		ELSE
				IF (_eDirection=E_Direction.DIRECTION_POSITIVE)THEN
					_fDistance:=_fPos-stAxis.stNcTOPLC.fActPos;
				ELSE
					_fDistance:=stAxis.stNcTOPLC.fActPos-_fPos;
				END_IF
		END_IF
		(*IF (_eDirection=E_Direction.DIRECTION_POSITIVE)THEN
			_fDistance:=_fPos-stAxis.stNcTOPLC.fActPos;
		ELSE
			_fDistance:=stAxis.stNcTOPLC.fActPos-_fPos;
		END_IF*)
		_nPathSegment:=1;
		_fAcc:=stAxis.stPLCTONC.stEndPosition.fAccleration;
	    _fDec:=stAxis.stPLCTONC.stEndPosition.fDeceleration;
ELSE
		_nPathSegment:=2;
		_fVeloStart:=stAxis.stNcTOPLC.fActVelo;
	    _fVeloEnd:=_fPreTaVel;
	    _fTargetVelo:=_fPreTaVel;
		_fDistance:=_fNewAccDis;
		_fAcc:=_fNewAcc;
	    _fDec:=_fNewAcc;
		_fPosIn:=_fDealt_S+_fPreDealt_S;       //11.29
	    _fVeloStart_2:=_fPreTaVel;
	    _fVeloEnd_2:=0.0;
	    _fTargetVelo_2:=_fPreTaVel;
		IF (stAxis.stPLCTONC.nRoadID_2<>0)AND (stAxis.stPLCTONC.nRoadID_1<>0)THEN   //判断指令
				IF (stAxis.stPLCTONC.stStartPosition.nRoadID<>stAxis.stPLCTONC.stEndPosition.nRoadID)THEN
				    IF(stAxis.stNcTOPLC.nCuRoadID=stAxis.stPLCTONC.nRoadID_2) THEN //第二路段
						IF (_eDirection=E_Direction.DIRECTION_POSITIVE)THEN
							 IF NOT stAxis.stPLCTONC.bRoadDirection  THEN   //正向 
								 _fDistance_2:=_fPos-stAxis.stPLCTONC.fRoad1_Length-stAxis.stNcTOPLC.fActPos-_fNewAccDis;
							 ELSE
								 _fDistance_2:=stAxis.stNcTOPLC.fActPos-(stAxis.stPLCTONC.fRoad2_Length-_fPos+stAxis.stPLCTONC.fRoad1_Length)-_fNewAccDis;
							 END_IF
						ELSE
							IF NOT stAxis.stPLCTONC.bRoadDirection  THEN   //正向 
								 _fDistance_2:=ABS(_fPos)-stAxis.stNcTOPLC.fActPos-_fNewAccDis;
							 ELSE
								 _fDistance_2:=stAxis.stNcTOPLC.fActPos-(stAxis.stPLCTONC.fRoad2_Length-ABS(_fPos))-_fNewAccDis;
							 END_IF
						END_IF
						stAxis.stPLCTONC.stStartPosition.nRoadID:=stAxis.stNcTOPLC.nCuRoadID;
					ELSE
						IF (_eDirection=E_Direction.DIRECTION_POSITIVE)THEN
							_fDistance_2:=_fPos-stAxis.stNcTOPLC.fActPos-_fNewAccDis;
						ELSE
							_fDistance_2:=stAxis.stNcTOPLC.fActPos-_fPos-_fNewAccDis;
						END_IF
					END_IF
				ELSE
					IF(stAxis.stNcTOPLC.nCuRoadID=stAxis.stPLCTONC.nRoadID_2) THEN //第二路段
						
						IF NOT stAxis.stPLCTONC.bRoadDirection  THEN   //正向 
							_fDistance_2:=_fPos-stAxis.stNcTOPLC.fActPos-_fNewAccDis;
						ELSE
							_fDistance_2:=stAxis.stNcTOPLC.fActPos-_fPos-_fNewAccDis;
						END_IF
						stAxis.stPLCTONC.stStartPosition.nRoadID:=stAxis.stNcTOPLC.nCuRoadID;
					ELSE
						IF (_eDirection=E_Direction.DIRECTION_POSITIVE)THEN
							_fDistance_2:=_fPos-stAxis.stNcTOPLC.fActPos-_fNewAccDis;
						ELSE
							_fDistance_2:=stAxis.stNcTOPLC.fActPos-_fPos-_fNewAccDis;
						END_IF
					END_IF
				END_IF
		ELSE
				IF (_eDirection=E_Direction.DIRECTION_POSITIVE)THEN
					_fDistance_2:=_fPos-stAxis.stNcTOPLC.fActPos-_fNewAccDis;
				ELSE
					_fDistance_2:=stAxis.stNcTOPLC.fActPos-_fPos-_fNewAccDis;
				END_IF
		END_IF
		(*IF (_eDirection=E_Direction.DIRECTION_POSITIVE)THEN
			_fDistance_2:=_fPos-stAxis.stNcTOPLC.fActPos-_fNewAccDis;
		ELSE
			_fDistance_2:=stAxis.stNcTOPLC.fActPos-_fPos-_fNewAccDis;
		END_IF*)
		_fAcc_2:=stAxis.stPLCTONC.stEndPosition.fAccleration;
	    _fDec_2:=stAxis.stPLCTONC.stEndPosition.fDeceleration;
		
END_IF
_bSynMode:=TRUE;
_bEnable:=TRUE;
stAxis.stAxisStatus.bSynDecActive:=TRUE;
IF GVL_MC.cDebug  THEN
	_sMessage:=FC_StrContact(stAxis,'next road dec2 gap control');
	 ADSLOGSTR(ADSLOG_MSGTYPE_HINT, _sMessage, '');
END_IF
END_ACTION

ACTION A_NextRoadGapControl:

//IF ((_fRealDis -_fGapSet)<=cDealtGap)AND(_pNextRoadPremover^.stAxisStatus.stPathRef.fTargetVelocity <stAxis.stAxisStatus.stPathRef.fTargetVelocity) THEN    //10.18 
(*IF ((_fRealDis -_fGapSet)<=_fSetDealtGap)AND(_pNextRoadPremover^.stAxisStatus.stPathRef.fTargetVelocity <stAxis.stAxisStatus.stPathRef.fTargetVelocity) THEN    //10.18
	
		_fPos:=stAxis.stPLCTONC.stEndPosition.fPosition;
		_fTargetVelo:=_pNextRoadPremover^.stAxisStatus.stPathRef.fTargetVelocity;
		_fVeloStart:=stAxis.stNcTOPLC.fActVelo;
		_fVeloEnd:=0;
		_fAcc:=stAxis.stPLCTONC.stEndPosition.fAccleration;
		_fDec:=stAxis.stPLCTONC.stEndPosition.fDeceleration;
		IF (_eDirection=E_Direction.DIRECTION_POSITIVE)THEN
		     _fDistance:=_fPos-stAxis.stNcTOPLC.fActPos;
	    ELSE
			 _fDistance:=stAxis.stNcTOPLC.fActPos-_fPos;
	    END_IF
		_bEnable:=TRUE;
		_nPathSegment:=1;
		stAxis.stAxisStatus.bSynDecActive:=TRUE;
		IF GVL_MC.cDebug  THEN
		     _sMessage:=FC_StrContact(stAxis,'nextroad gap control');
	         ADSLOGSTR(ADSLOG_MSGTYPE_HINT, _sMessage, '');
        END_IF
		RETURN;
END_IF *)

IF _fRealDis <=0 THEN   //05.19
	RETURN;
END_IF

IF (_pNextRoadPremover^.stAxisStatus.nNcCycleCounter<>0)THEN 
	 A_NextRoadCatchUp();
   // IF ((_fRealDis -_fGapSet)<=cDealtGap) THEN    //10.18 
	IF ((_fRealDis -_fGapSet)<=_fSetDealtGap) THEN    //10.18 	
			IF _fbDecNextPathTrig.Q THEN 
					   IF (stAxis.stPLCTONC.nRoadID_2<>0)AND (stAxis.stPLCTONC.nRoadID_1<>0)AND(stAxis.stNcTOPLC.nCuRoadID=stAxis.stPLCTONC.nRoadID_2)THEN
						   IF (stAxis.stPLCTONC.stStartPosition.nRoadID<>stAxis.stPLCTONC.stEndPosition.nRoadID)THEN
								IF (_eDirection=E_Direction.DIRECTION_POSITIVE)THEN
									IF NOT stAxis.stPLCTONC.bRoadDirection  THEN
										 _fPos:=stAxis.stPLCTONC.stEndPosition.fPosition-stAxis.stPLCTONC.fRoad1_Length;
									ELSE
										_fPos:=stAxis.stPLCTONC.fRoad2_Length-(stAxis.stPLCTONC.stEndPosition.fPosition-stAxis.stPLCTONC.fRoad1_Length);
									END_IF
									_fDistance:=ABS(stAxis.stNcTOPLC.fActPos-_fPos);
								ELSE
									IF NOT stAxis.stPLCTONC.bRoadDirection  THEN
										 _fPos:=ABS(stAxis.stPLCTONC.stEndPosition.fPosition);
									ELSE
										_fPos:=stAxis.stPLCTONC.fRoad2_Length-ABS(stAxis.stPLCTONC.stEndPosition.fPosition);
									END_IF
									_fDistance:=ABS(stAxis.stNcTOPLC.fActPos-_fPos);
								END_IF
						   ELSE
								_fPos:=stAxis.stPLCTONC.stEndPosition.fPosition;
								_fDistance:=ABS(stAxis.stNcTOPLC.fActPos-_fPos);
						   END_IF
					   ELSE
						   _fPos:=stAxis.stPLCTONC.stEndPosition.fPosition;
						   IF (_eDirection=E_Direction.DIRECTION_POSITIVE)THEN
							  _fDistance:=_fPos-stAxis.stNcTOPLC.fActPos;
						   ELSE
							  _fDistance:=stAxis.stNcTOPLC.fActPos-_fPos;
						   END_IF
					   END_IF
					   //_fPos:=stAxis.stPLCTONC.stEndPosition.fPosition;
					   IF _pNextRoadPremover^.stPLCTONC.bCmdDceUpdate THEN
							_fTargetVelo:=_pNextRoadPremover^.stPLCTONC.fTargetVelocity;
					   ELSE
						   _fTargetVelo:=_pNextRoadPremover^.stAxisStatus.stPathRef.fTargetVelocity;
					   END_IF
					   //_fTargetVelo:=_pNextRoadPremover^.stAxisStatus.stPathRef.fTargetVelocity;
					   _fVeloStart:=stAxis.stNcTOPLC.fActVelo;
					   _fVeloEnd:=0;
					   _fAcc:=stAxis.stPLCTONC.stEndPosition.fAccleration;
					   _fDec:=stAxis.stPLCTONC.stEndPosition.fDeceleration;
					   
					   _bEnable:=TRUE;
					   _nPathSegment:=1;
					   stAxis.stAxisStatus.bSynDecActive:=TRUE;
					   IF GVL_MC.cDebug  THEN
						_sMessage:=FC_StrContact(stAxis,'Nextroad SynDecActive path');
						 ADSLOGSTR(ADSLOG_MSGTYPE_HINT, _sMessage, '');
					   END_IF
			END_IF
	END_IF

END_IF
END_ACTION

ACTION A_NodeConfig:
IF stAxis.stNcTOPLC.nCuRoadID=0 THEN 
	RETURN;
END_IF 

_nMoverCounter:=GVL_MC.aRoadRef[stAxis.stNcTOPLC.nCuRoadID].nMoverCounter;
IF _nMoverCounter<>_nLastMoverCounter AND _nMoverCounter<>0  THEN 
	
    FOR _nNodeIndex:=1 TO GVL_MC.MAX_MOVER  DO
	    IF (GVL_MC.aRoadRef[stAxis.stNcTOPLC.nCuRoadID].aNode[_nNodeIndex].nAxisId=stAxis.stNcTOPLC.nAxisId)THEN
			stAxis.stAxisStatus.pPremover:=GVL_MC.aRoadRef[stAxis.stNcTOPLC.nCuRoadID].aNode[_nNodeIndex].pPremover;
	        stAxis.stAxisStatus.pAftermover:=GVL_MC.aRoadRef[stAxis.stNcTOPLC.nCuRoadID].aNode[_nNodeIndex].pAftermover;
			EXIT;
		END_IF
   END_FOR
   _nLastMoverCounter:=GVL_MC.aRoadRef[stAxis.stNcTOPLC.nCuRoadID].nMoverCounter;   //05.08 修改前置后置更新条件
END_IF
END_ACTION

ACTION A_NodeUpdate:
// road node 更新
// 动子出现在某road上增加 01.09
_fbTrigRoadUpdate(CLK:=stAxis.stCodToNCParam.bArrayReseved1 , Q=> );
//IF stAxis.stNcTOPLC.nCuRoadID=0 AND stAxis.stCodToNCParam.bArrayReseved1  AND stAxis.stCodToNCParam.nRoadID<>0 THEN
IF _fbTrigRoadUpdate.Q  AND stAxis.stCodToNCParam.nRoadID<>0 AND NOT _bInsertOk THEN
	stAxis.stNcTOPLC.nCuRoadID:=stAxis.stCodToNCParam.nRoadID;
	_bInsertOk :=_fbAxisGroupList.M_InsertNode(aRoadRef:=GVL_MC.aRoadRef , nSysType:=stAxis.stAxisParam.stRoadParam.nSysType , nRoadId:=stAxis.stCodToNCParam.nRoadID , pAixs:=ADR(stAxis) );
    (*IF GVL_MC.cDebug  THEN
	    _sMessage2:=FC_StrContactEx(stAxis,'insertAxis');
	     ADSLOGSTR(ADSLOG_MSGTYPE_HINT, _sMessage2, '');
    END_IF*)
	_sMessage3:='';
	_sMessage3:=CONCAT(DWORD_TO_STRING(stAxis.stNcTOPLC.nAxisId),',insertAxis');
	IF stAxis.stNcTOPLC.nCuRoadID>0 AND stAxis.stNcTOPLC.nCuRoadID<=GVL_MC.cRoadNum AND GVL_MC.cDebug THEN
		IF GVL_MC.aRoadRef[stAxis.stNcTOPLC.nCuRoadID].nMoverCounter>0  THEN
			FOR _nPreIndex:=1 TO GVL_MC.aRoadRef[stAxis.stNcTOPLC.nCuRoadID].nMoverCounter   DO
				_sMessage3:=CONCAT(_sMessage3,DWORD_TO_STRING(GVL_MC.aRoadRef[stAxis.stNcTOPLC.nCuRoadID].aNode[_nPreIndex].nAxisId));
				_sMessage3:=CONCAT(_sMessage3,',');
			END_FOR
			ADSLOGSTR(ADSLOG_MSGTYPE_HINT, _sMessage3, '');
		END_IF
	END_IF
END_IF
IF NOT stAxis.stCodToNCParam.bArrayReseved1 THEN
	_bInsertOk:=FALSE;
END_IF
// 07.04
IF stAxis.stNcTOPLC.nCuRoadID=0 THEN 
	RETURN;
END_IF 

_fbTrigRoadDeleUpdate(CLK:=stAxis.stCodToNCParam.bArrayReseved2 , Q=> );   //01.29
IF _fbTrigRoadDeleUpdate.Q THEN
	_bDeleteNodeOk:=_fbAxisGroupList.M_DeleteNode(aRoadRef:=GVL_MC.aRoadRef , nSysType:=stAxis.stAxisParam.stRoadParam.nSysType , nRoadId:=stAxis.stNcTOPLC.nCuRoadID , pAixs:=ADR(stAxis));
	(*IF GVL_MC.cDebug  THEN
	    _sMessage2:=FC_StrContactEx(stAxis,'deleteAxis');
	     ADSLOGSTR(ADSLOG_MSGTYPE_HINT, _sMessage2, '');
    END_IF*)
	_sMessage3:='';
	_sMessage3:=CONCAT(DWORD_TO_STRING(stAxis.stNcTOPLC.nAxisId),',deleteAxis');
    IF stAxis.stNcTOPLC.nCuRoadID>0 AND stAxis.stNcTOPLC.nCuRoadID<=GVL_MC.cRoadNum AND GVL_MC.cDebug THEN
	    IF GVL_MC.aRoadRef[stAxis.stNcTOPLC.nCuRoadID].nMoverCounter>0 THEN
			FOR _nPreIndex:=1 TO GVL_MC.aRoadRef[stAxis.stNcTOPLC.nCuRoadID].nMoverCounter   DO
				_sMessage3:=CONCAT(_sMessage3,DWORD_TO_STRING(GVL_MC.aRoadRef[stAxis.stNcTOPLC.nCuRoadID].aNode[_nPreIndex].nAxisId));
				_sMessage3:=CONCAT(_sMessage3,',');
			END_FOR
			ADSLOGSTR(ADSLOG_MSGTYPE_HINT, _sMessage3, '');
		END_IF
	END_IF
END_IF

// 先增加后删除
(*IF stAxis.stNcTOPLC.nCuRoadID=0 THEN 
	RETURN;
END_IF *) //07.04
IF (_nLastRoadID<>stAxis.stNcTOPLC.nCuRoadID) AND (_nLastRoadID<>0)THEN
	
	_nLastMoverCounter:=GVL_MC.aRoadRef[stAxis.stNcTOPLC.nCuRoadID].nMoverCounter;  //********重新修改前置后质更新条件     05.08
	_bAddNodeOk :=_fbAxisGroupList.M_AddNode(aRoadRef:=GVL_MC.aRoadRef , nRoadId:=stAxis.stNcTOPLC.nCuRoadID , pAixs:=ADR(stAxis));
	//_bAddNodeOk :=_fbAxisGroupList.M_InsertNode(aRoadRef:=GVL_MC.aRoadRef , nSysType:=stAxis.stAxisParam.stRoadParam.nSysType , nRoadId:=stAxis.stNcTOPLC.nCuRoadID , pAixs:=ADR(stAxis) );
    _bDeleteNodeOk:=_fbAxisGroupList.M_DeleteNode(aRoadRef:=GVL_MC.aRoadRef , nSysType:=stAxis.stAxisParam.stRoadParam.nSysType , nRoadId:=_nLastRoadID , pAixs:=ADR(stAxis));
	(*IF GVL_MC.cDebug  THEN
	    //_sMessage2:=FC_StrContactEx(stAxis,'roadchange');
	    // ADSLOGSTR(ADSLOG_MSGTYPE_HINT, _sMessage2, '');
		  _sMessage3:=CONCAT(DWORD_TO_STRING(stAxis.stNcTOPLC.nAxisId),',roadchange');
		  _sMessage3:=CONCAT(_sMessage3,',');
		  _sMessage3:=CONCAT(_sMessage3,LREAL_TO_STRING(stAxis.stNcTOPLC.fActPos));
		  _sMessage3:=CONCAT(_sMessage3,',');
		  _sMessage3:=CONCAT(_sMessage3,DWORD_TO_STRING(GVL_MC.aRoadRef[stAxis.stNcTOPLC.nCuRoadID].aNode[GVL_MC.aRoadRef[stAxis.stNcTOPLC.nCuRoadID].nMoverCounter].pMover^.stNcTOPLC.nAxisId));
          _sMessage3:=CONCAT(_sMessage3,',');	 
		  _sMessage3:=CONCAT(_sMessage3,LREAL_TO_STRING(GVL_MC.aRoadRef[stAxis.stNcTOPLC.nCuRoadID].aNode[GVL_MC.aRoadRef[stAxis.stNcTOPLC.nCuRoadID].nMoverCounter].pMover^.stNcTOPLC.fActPos));
   	      _sMessage3:=CONCAT(_sMessage3,',');
		  _sMessage3:=CONCAT(_sMessage3,UINT_TO_STRING(GVL_MC.aRoadRef[stAxis.stNcTOPLC.nCuRoadID].nMoverCounter));
		  ADSLOGSTR(ADSLOG_MSGTYPE_HINT, _sMessage3, '');
    END_IF*)
	_sMessage3:='';
	_sMessage3:=CONCAT(DWORD_TO_STRING(stAxis.stNcTOPLC.nAxisId),',roadchange');
	IF stAxis.stNcTOPLC.nCuRoadID>0 AND stAxis.stNcTOPLC.nCuRoadID<=GVL_MC.cRoadNum AND GVL_MC.cDebug THEN
		IF GVL_MC.aRoadRef[stAxis.stNcTOPLC.nCuRoadID].nMoverCounter>0  THEN
			FOR _nPreIndex:=1 TO GVL_MC.aRoadRef[stAxis.stNcTOPLC.nCuRoadID].nMoverCounter   DO
				
				_sMessage3:=CONCAT(_sMessage3,DWORD_TO_STRING(GVL_MC.aRoadRef[stAxis.stNcTOPLC.nCuRoadID].aNode[_nPreIndex].nAxisId));
				_sMessage3:=CONCAT(_sMessage3,',');
			END_FOR
			ADSLOGSTR(ADSLOG_MSGTYPE_HINT, _sMessage3, '');
		END_IF
	END_IF
END_IF



_nLastRoadID:=stAxis.stNcTOPLC.nCuRoadID;

_bAddNodeOk:=FALSE;
_bDeleteNodeOk:=FALSE;
END_ACTION

ACTION A_Planning:
IF (stAxis.stPLCTONC.ePlanningMode=E_PlanningMode.PLANNINGMODE_TSHAPED)THEN 
   A_TShaped();
ELSIF (stAxis.stPLCTONC.ePlanningMode=E_PlanningMode.PLANNINGMODE_SSHAPED)THEN 
   A_SShapedPlanning();
ELSIF (stAxis.stPLCTONC.ePlanningMode=E_PlanningMode.PLANNINGMODE_LINEAR)THEN 
  A_LinearPlanning();

ELSIF (stAxis.stPLCTONC.ePlanningMode=E_PlanningMode.PLANNINGMODE_FOLLOWMASTER)THEN 
  A_FollowMasterPlanning();
  
ELSIF (stAxis.stPLCTONC.ePlanningMode=E_PlanningMode.PLANNINGMODE_PLOYNOM3)THEN 
	A_Ploynom3Planning();
ELSIF (stAxis.stPLCTONC.ePlanningMode=E_PlanningMode.PLANNINGMODE_FOLLOW)THEN 
	A_FollowPlanning();	
ELSE 
   A_TShaped();

END_IF
END_ACTION

ACTION A_Ploynom3Planning:
//_fbAxis.strStartPoint.fPosition:=stAxis.stNcTOPLC.fActPos;
//_fbAxis.strEndPoint.fPosition:=stAxis.stPLCTONC.stEndPosition.fPosition;
_fbAxis.strStartPoint.fPosition:=0;
_fbAxis.strEndPoint.fPosition:=ABS(stAxis.stPLCTONC.stEndPosition.fPosition-stAxis.stNcTOPLC.fActPos)/ABS(stAxis.stPLCTONC.stMasterParam.fEndPos-stAxis.stPLCTONC.stMasterParam.fStartPos);

IF (stAxis.stAxisStatus.pMaster^.stNcTOPLC.fActVelo<>0)  THEN 
    _fbAxis.strStartPoint.fVelocity :=stAxis.stNcTOPLC.fActVelo/stAxis.stAxisStatus.pMaster^.stNcTOPLC.fActVelo;
ELSE
	_fbAxis.strStartPoint.fVelocity :=0;
END_IF

//_fbAxis.strEndPoint.fVelocity:=stAxis.stAxisStatus.stPathRef.fVeloRatio;
_fbAxis.strEndPoint.fVelocity:=stAxis.stPLCTONC.fGearRatio;
_stPolynom5Factor:=_fbAxis.M_Ploynom3(fTheat_Start:=0 ,
               fTheat_End:=1  );
			   

_bCalculateDone:=TRUE;
END_ACTION

ACTION A_Ploynom3Position:
_nSysType:=stAxis.stPLCTONC.nSysType;
stAxis.stNcTOPLC.nAxisState:=6;
stAxis.stAxisStatus.nNcCycleCounter:=stAxis.stAxisStatus.nNcCycleCounter+1;
_fMasterStartPos:=stAxis.stPLCTONC.stMasterParam.fStartPos;
_fMasterEndPos:=stAxis.stPLCTONC.stMasterParam.fEndPos;

_fSlaveStartPos:=stAxis.stPLCTONC.stStartPosition.fPosition;
// 自变量区间归一化

_fDealt_X:=ABS(_fMasterEndPos-_fMasterStartPos);
IF (_fDealt_X<=0)THEN 
	RETURN;
END_IF
_fPos_X:=ABS(stAxis.stAxisStatus.pMaster^.stNcTOPLC.fActPos-_fMasterStartPos)/_fDealt_X;

IF (_fPos_X<=1)THEN

	// 归一化从轴位置、速度、加速度和加加速计算
	_stAxis_Point.fPosition:=_stPolynom5Factor.fA0+ _stPolynom5Factor.fA1*_fPos_X+ _stPolynom5Factor.fA2*_fPos_X*_fPos_X
						   +_stPolynom5Factor.fA3*_fPos_X*_fPos_X*_fPos_X; 
						   
	_stAxis_Point.fVelocity:=_stPolynom5Factor.fA1+ 2*_stPolynom5Factor.fA2*_fPos_X+3*_stPolynom5Factor.fA3*_fPos_X*_fPos_X;
	
	_stAxis_Point.fAccleration:=2*_stPolynom5Factor.fA2+6*_stPolynom5Factor.fA3*_fPos_X;
	_stAxis_Point.fbJerk:=6*_stPolynom5Factor.fA3;
	
	IF stAxis.stAxisStatus.bPositiveDirection THEN
		stAxis.stNcTOPLC.fActPos:=_fDealt_X*_stAxis_Point.fPosition+_fSlaveStartPos;    
	ELSE
		stAxis.stNcTOPLC.fActPos:=_fSlaveStartPos-_fDealt_X*_stAxis_Point.fPosition;    
	END_IF                  
	stAxis.stNcTOPLC.fSetVelo:=_stAxis_Point.fVelocity*ABS(stAxis.stAxisStatus.pMaster^.stNcTOPLC.fActVelo);
	stAxis.stNcTOPLC.fSetAcc:=_stAxis_Point.fAccleration*ABS(stAxis.stAxisStatus.pMaster^.stNcTOPLC.fActVelo*stAxis.stAxisStatus.pMaster^.stNcTOPLC.fActVelo)/_fDealt_X;
	stAxis.stNcTOPLC.fSetJerk:=_stAxis_Point.fbJerk*ABS(stAxis.stAxisStatus.pMaster^.stNcTOPLC.fActVelo*stAxis.stAxisStatus.pMaster^.stNcTOPLC.fActVelo*stAxis.stAxisStatus.pMaster^.stNcTOPLC.fActVelo)/(_fDealt_X*_fDealt_X);
							  
	stAxis.stNcTOPLC.fActVelo:=stAxis.stNcTOPLC.fSetVelo;
	_stAxis_Point.fPosition:=stAxis.stNcTOPLC.fActPos;
ELSE
	stAxis.stNcTOPLC.fSetVelo:=LTRUNC(stAxis.stAxisStatus.pMaster^.stNcTOPLC.fActVelo*stAxis.stPLCTONC.fGearRatio);
    stAxis.stNcTOPLC.fActVelo:=LTRUNC(stAxis.stAxisStatus.pMaster^.stNcTOPLC.fActVelo*stAxis.stPLCTONC.fGearRatio);
    IF stAxis.stAxisStatus.bPositiveDirection THEN
         _stAxis_Point.fPosition:=stAxis.stAxisStatus.pMaster^.stNcTOPLC.fDealtPos*stAxis.stPLCTONC.fGearRatio +_stAxis_Point.fPosition;

    ELSE
        _stAxis_Point.fPosition:=-stAxis.stAxisStatus.pMaster^.stNcTOPLC.fDealtPos*stAxis.stPLCTONC.fGearRatio +_stAxis_Point.fPosition;
    END_IF
	stAxis.stNcTOPLC.fDealtPos:=ABS(LTRUNC(_stAxis_Point.fPosition)-stAxis.stNcTOPLC.fActPos);    //01.13
	stAxis.stNcTOPLC.fActPos:=LTRUNC(_stAxis_Point.fPosition);
END_IF
END_ACTION

ACTION A_Ploynom5Position:
_bEndOfProfile:=FALSE;
_nSysType:=stAxis.stPLCTONC.nSysType;
stAxis.stNcTOPLC.nAxisState:=6;
stAxis.stAxisStatus.nNcCycleCounter:=stAxis.stAxisStatus.nNcCycleCounter+1;

//数据装载
IF stAxis.stPLCTONC.stCamParam.bCamLoad THEN 
   _stCamParam:=stAxis.stPLCTONC.stCamParam;
   stAxis.stPLCTONC.stCamParam.bCamLoad:=FALSE;
END_IF 

//buffer 更新
 _fbCamBufUpdateTrig(CLK:= (INT_TO_UINT(_nIndex)=(cPointBuffer-1)OR (NOT _bFisrtUpdate)), Q=> );

IF(_stCamParam.nElements> cPointBuffer) THEN
   IF _fbCamBufUpdateTrig.Q   THEN
      _aCamBuffer:=_stCamParam.aCamBuffer;
	  _nIndex:=0;
	  _nCamBufferNum:=_nCamBufferNum+1;
   END_IF 
ELSE
	_aCamBuffer:=_stCamParam.aCamBuffer;
	_nCamBufferNum:=1;
END_IF

// 点更新及曲线系数计算
_fbCamPointUpdateTrig(CLK:=(_nIndex<>_nLastIndex)OR (NOT _bFisrtUpdate)   , Q=> );
IF _fbCamPointUpdateTrig.Q THEN
     IF (_stCamParam.nPointType=1) THEN  //xyva
         _fMasterStartPos:=_aCamBuffer[_nIndex].fDx;
	     _fMasterEndPos:=_aCamBuffer[_nIndex+1].fDx;
	     _fDealt_X:=ABS(_fMasterEndPos-_fMasterStartPos);
		 IF (_fDealt_X=0)THEN 
			 RETURN;
		 END_IF
		_fSlaveStartPos :=_aCamBuffer[_nIndex].fDy;
		_fbAxis.strStartPoint.fPosition:=0;
		_fbAxis.strEndPoint.fPosition:=ABS((_aCamBuffer[_nIndex+1].fDy-_fSlaveStartPos))/_fDealt_X;
		_fbAxis.strStartPoint.fVelocity :=_aCamBuffer[_nIndex].fDv;
		_fbAxis.strEndPoint.fVelocity:=_aCamBuffer[_nIndex+1].fDv;
		_fbAxis.strStartPoint.fAccleration :=_aCamBuffer[_nIndex].fDa*_fDealt_X;
		_fbAxis.strEndPoint.fAccleration:=_aCamBuffer[_nIndex+1].fDa*_fDealt_X;
		_fbAxis.strStartPoint.fbJerk :=_aCamBuffer[_nIndex].fDa*_fDealt_X*_fDealt_X;
		_fbAxis.strEndPoint.fbJerk:=_aCamBuffer[_nIndex+1].fDa*_fDealt_X*_fDealt_X;
	 ELSIF (_stCamParam.nPointType=2) THEN   //xy
		 _fMasterStartPos:=_aCamBuffer[_nIndex].fDx;
	     _fMasterEndPos:=_aCamBuffer[_nIndex+1].fDx;
	     _fDealt_X:=ABS(_fMasterEndPos-_fMasterStartPos);
		 _fSlaveStartPos :=_aCamBuffer[_nIndex].fDy;
		 _fbAxis.strStartPoint.fPosition:=0;
		 IF (_fDealt_X=0)THEN 
			 RETURN;
		 END_IF
		 _fbAxis.strEndPoint.fPosition:=ABS(_aCamBuffer[_nIndex+1].fDy-_fSlaveStartPos)/_fDealt_X;
		 IF (_nIndex=0)AND (_nCamBufferNum=1)THEN
		    _fbAxis.strStartPoint.fVelocity :=0;
			_fbAxis.strStartPoint.fAccleration :=0;
		 ELSE
			 _fbAxis.strStartPoint.fVelocity :=1;
			 _fbAxis.strStartPoint.fAccleration :=0;
		 END_IF

		 _fbAxis.strEndPoint.fVelocity:=1;
		 IF _stCamParam.bPeriodic AND (stAxis.stNcTOPLC.nCuSegIndex =(_stCamParam.nElements-1)) THEN
			 _fbAxis.strEndPoint.fVelocity:=0;
		 END_IF
		 _fbAxis.strStartPoint.fAccleration :=0;
		 _fbAxis.strEndPoint.fAccleration:=0;
		 _fbAxis.strStartPoint.fbJerk :=0;
		 _fbAxis.strEndPoint.fbJerk:=0;
		
     ELSE
		 RETURN;
		 
	 END_IF
	_stPolynom5Factor:=_fbAxis.M_Ploynom5(fTheat_Start:=0 ,fTheat_End:=1);
	_bFisrtUpdate:=TRUE;
END_IF 
_nLastIndex :=_nIndex;
IF (_fDealt_X=0)THEN 
	RETURN;
END_IF
// 位置计算

// 自变量区间归一化
//_fDealt_X:=_fMasterEndPos-_fMasterStartPos;
IF stAxis.stAxisStatus.bPositiveDirection  THEN
    _fPos_X:=(stAxis.stAxisStatus.pMaster^.stNcTOPLC.fActPos-_fMasterStartPos)/ABS(_fDealt_X);
ELSE
	_fPos_X:=(_fMasterStartPos-stAxis.stAxisStatus.pMaster^.stNcTOPLC.fActPos)/ABS(_fDealt_X);
END_IF

IF (_fPos_X<0)THEN 
	RETURN;
END_IF

_stAxis_Point.fPosition:=_stPolynom5Factor.fA0+ _stPolynom5Factor.fA1*_fPos_X+ _stPolynom5Factor.fA2*_fPos_X*_fPos_X
                        +_stPolynom5Factor.fA3*_fPos_X*_fPos_X*_fPos_X+_stPolynom5Factor.fA4*_fPos_X*_fPos_X*_fPos_X*_fPos_X
						+_stPolynom5Factor.fA5*_fPos_X*_fPos_X*_fPos_X*_fPos_X*_fPos_X;
                          
						
_stAxis_Point.fVelocity:=_stPolynom5Factor.fA1+ 2*_stPolynom5Factor.fA2*_fPos_X+3*_stPolynom5Factor.fA3*_fPos_X*_fPos_X
                          +4*_stPolynom5Factor.fA4*_fPos_X*_fPos_X*_fPos_X+5*_stPolynom5Factor.fA5*_fPos_X*_fPos_X*_fPos_X*_fPos_X;
                          
_stAxis_Point.fAccleration:= 2*_stPolynom5Factor.fA2+6*_stPolynom5Factor.fA3*_fPos_X+12*_stPolynom5Factor.fA4*_fPos_X*_fPos_X+20*_stPolynom5Factor.fA5*_fPos_X*_fPos_X*_fPos_X;
_stAxis_Point.fbJerk:=6*_stPolynom5Factor.fA3+24*_stPolynom5Factor.fA4*_fPos_X+60*_stPolynom5Factor.fA5*_fPos_X*_fPos_X;

IF stAxis.stAxisStatus.bPositiveDirection THEN 
	//stAxis.stNcTOPLC.fSetPos:=_stAxis_Point.fPosition*_fDealt_X+_fSlaveStartPos;
	stAxis.stNcTOPLC.fActPos:=_stAxis_Point.fPosition*_fDealt_X+_fSlaveStartPos;
	stAxis.stNcTOPLC.fSetVelo:=_stAxis_Point.fVelocity*ABS(stAxis.stAxisStatus.pMaster^.stNcTOPLC.fActVelo);
	stAxis.stNcTOPLC.fSetAcc:=_stAxis_Point.fAccleration*ABS(stAxis.stAxisStatus.pMaster^.stNcTOPLC.fActVelo*stAxis.stAxisStatus.pMaster^.stNcTOPLC.fActVelo)/_fDealt_X;
	stAxis.stNcTOPLC.fSetJerk:=_stAxis_Point.fbJerk*ABS(stAxis.stAxisStatus.pMaster^.stNcTOPLC.fActVelo*stAxis.stAxisStatus.pMaster^.stNcTOPLC.fActVelo*stAxis.stAxisStatus.pMaster^.stNcTOPLC.fActVelo)/(_fDealt_X*_fDealt_X);
	//stAxis.stNcTOPLC.fActPos:=stAxis.stNcTOPLC.fSetPos;
	stAxis.stNcTOPLC.fActVelo:=stAxis.stNcTOPLC.fSetVelo;
ELSE
	//stAxis.stNcTOPLC.fSetPos:=-_stAxis_Point.fPosition*_fDealt_X+_fSlaveStartPos;
	stAxis.stNcTOPLC.fActPos:=-_stAxis_Point.fPosition*_fDealt_X+_fSlaveStartPos;
	stAxis.stNcTOPLC.fSetVelo:=_stAxis_Point.fVelocity*ABS(stAxis.stAxisStatus.pMaster^.stNcTOPLC.fActVelo);
	stAxis.stNcTOPLC.fSetAcc:=_stAxis_Point.fAccleration*ABS(stAxis.stAxisStatus.pMaster^.stNcTOPLC.fActVelo*stAxis.stAxisStatus.pMaster^.stNcTOPLC.fActVelo)/_fDealt_X;
	stAxis.stNcTOPLC.fSetJerk:=_stAxis_Point.fbJerk*ABS(stAxis.stAxisStatus.pMaster^.stNcTOPLC.fActVelo*stAxis.stAxisStatus.pMaster^.stNcTOPLC.fActVelo*stAxis.stAxisStatus.pMaster^.stNcTOPLC.fActVelo)/(_fDealt_X*_fDealt_X);
	//stAxis.stNcTOPLC.fActPos:=stAxis.stNcTOPLC.fSetPos;
	stAxis.stNcTOPLC.fActVelo:=stAxis.stNcTOPLC.fSetVelo;
END_IF
(*IF (_nSysType=3)THEN   //环形
	IF stAxis.stAxisStatus.bPositiveDirection THEN
		stAxis.stNcTOPLC.nModuloSetTurns:=LREAL_TO_DINT(LTRUNC(stAxis.stNcTOPLC.fSetPos/stAxis.stNcTOPLC.fModuloFactor));
	ELSE
		IF stAxis.stNcTOPLC.fSetPos<(stAxis.stNcTOPLC.nModuloSetTurns*stAxis.stNcTOPLC.fModuloFactor)THEN 
				stAxis.stNcTOPLC.nModuloSetTurns:=stAxis.stNcTOPLC.nModuloSetTurns-1;
		END_IF
	END_IF
	stAxis.stNcTOPLC.fModuloSetPos:= MODABS(stAxis.stNcTOPLC.fSetPos,stAxis.stNcTOPLC.fModuloFactor);
ELSE
	stAxis.stNcTOPLC.fModuloSetPos:= ABS(stAxis.stNcTOPLC.fSetPos);
END_IF*)


stAxis.stNcTOPLC.nCuSegIndex:=INT_TO_UINT(_nIndex+1)+(_nCamBufferNum-1)*cPointBuffer;
// index更新
IF stAxis.stAxisStatus.bPositiveDirection THEN 
	IF (stAxis.stNcTOPLC.fActPos>=_aCamBuffer[_nIndex+1].fDy)THEN 
		_nIndex:=_nIndex+1;
		IF stAxis.stNcTOPLC.nCuSegIndex >(_stCamParam.nElements-1) THEN      //结束条件判断
			_bCalculateDone:=FALSE;
			_nIndex:=0;
			_nLastIndex :=0;
			 stAxis.stAxisStatus.stPathRef.bCalculateDone:=FALSE;
			 stAxis.stNcTOPLC.nAxisState:=2;
		 
			 stAxis.stNcTOPLC.fSetAcc:=0;
			 _bFisrtUpdate:=FALSE;
			 stAxis.stNcTOPLC.nCuSegIndex:=0;
			 _nCamBufferNum:=0;
			 _fDealt_X:=0;
			 _fbCamBufUpdateTrig(CLK:= FALSE, Q=> );
			 _fbCamPointUpdateTrig(CLK:=FALSE   , Q=> );
			 _bEndOfProfile:=TRUE;
		END_IF
	END_IF
ELSE
	IF (stAxis.stNcTOPLC.fActPos<=_aCamBuffer[_nIndex+1].fDy)THEN 
		_nIndex:=_nIndex+1;
		IF stAxis.stNcTOPLC.nCuSegIndex >(_stCamParam.nElements-1) THEN      //结束条件判断
			_bCalculateDone:=FALSE;
			_nIndex:=0;
			_nLastIndex :=0;
			 stAxis.stAxisStatus.stPathRef.bCalculateDone:=FALSE;
			 stAxis.stNcTOPLC.nAxisState:=2;
		 
			 stAxis.stNcTOPLC.fSetAcc:=0;
			 _bFisrtUpdate:=FALSE;
			 stAxis.stNcTOPLC.nCuSegIndex:=0;
			 _nCamBufferNum:=0;
			 _fDealt_X:=0;
			 _fbCamBufUpdateTrig(CLK:= FALSE, Q=> );
			 _fbCamPointUpdateTrig(CLK:=FALSE   , Q=> );
			 _bEndOfProfile:=TRUE;
		END_IF
	END_IF
END_IF
END_ACTION

ACTION A_PositionHandle:
//stAxis.stNcTOPLC.fActPos 输入
//stAxis.stNcTOPLC.fSetPos输出
IF (stAxis.stPLCTONC.eCommand=E_Command.COMMAND_ABSOLUTEFORK)OR (stAxis.stPLCTONC.eCommand=E_Command.COMMAND_CAMIN)OR 
	(stAxis.stPLCTONC.eCommand=E_Command.COMMAND_GEARINPOS)THEN
	stAxis.stNcTOPLC.fSetPos:=stAxis.stNcTOPLC.fActPos;
    
ELSE
	IF (stAxis.stAxisParam.stRoadParam.nSysType=1) OR (stAxis.stAxisParam.stRoadParam.nSysType=4) THEN 
		stAxis.stNcTOPLC.fSetPos:=stAxis.stNcTOPLC.fActPos;
	ELSE
		_fbFilterV2(nWindowSize:=nWindowSize , fData:=stAxis.stNcTOPLC.fActPos , fOutputData=>stAxis.stNcTOPLC.fSetPos );
	END_IF
END_IF

IF (stAxis.stPLCTONC.nSysType=3)THEN
	IF stAxis.stAxisStatus.bPositiveDirection THEN
		stAxis.stNcTOPLC.nModuloSetTurns:=LREAL_TO_DINT(LTRUNC(stAxis.stNcTOPLC.fActPos/stAxis.stNcTOPLC.fModuloFactor));
	ELSE
		IF stAxis.stNcTOPLC.fActPos<(stAxis.stNcTOPLC.nModuloSetTurns*stAxis.stNcTOPLC.fModuloFactor)THEN 
			 stAxis.stNcTOPLC.nModuloSetTurns:=stAxis.stNcTOPLC.nModuloSetTurns-1;
		END_IF
	END_IF
							
	stAxis.stNcTOPLC.fModuloSetPos:= MODABS(stAxis.stNcTOPLC.fSetPos,stAxis.stNcTOPLC.fModuloFactor);
ELSE
	stAxis.stNcTOPLC.fModuloSetPos:=ABS(stAxis.stNcTOPLC.fSetPos);
	// 04.30增加环形位置同步
	IF (stAxis.stAxisParam.stRoadParam.nSysType=3)THEN
		stAxis.stNcTOPLC.fModuloSetPos:= MODABS(stAxis.stNcTOPLC.fSetPos,stAxis.stNcTOPLC.fModuloFactor);
	END_IF
END_IF
END_ACTION

ACTION A_SShapedPlanning:
_stSShapedParam:=_fbAxis.M_SShaped(
					fStartPos:=_fStartPos , 
					fEndPos:=_fEndPos , 
					fStartVelo:=_fVeloStart , 
					fEndVelo:=_fVeloEnd , 
					fTargetVelo:=_fTargetVelo , 
					fTargetAcc:=_fAcc , 
					fTargetJerk:=_fJerk );
					
_stPathRef._nPathSegmentNum:=1;
_stPathRef.aExecutablePath[0].fTa:=_stSShapedParam.fTa;
_stPathRef.aExecutablePath[0].fTv:=_stSShapedParam.fTv;
_stPathRef.aExecutablePath[0].fTd:=_stSShapedParam.fTd;
_stPathRef.aExecutablePath[0].fTj1:=_stSShapedParam.fTj1;
_stPathRef.aExecutablePath[0].fTj2:=_stSShapedParam.fTj2;
_stPathRef.aExecutablePath[0].fTotalTime:=_stSShapedParam.fT;


_stPathRef.aExecutablePath[0].fStartVelo:=_fVeloStart;
_stPathRef.aExecutablePath[0].fExpVelo:=_stSShapedParam.fVlim;
_stPathRef.aExecutablePath[0].fEndVelo:=_fVeloEnd;
_stPathRef.aExecutablePath[0].fAccleration:=_stSShapedParam.fA_LimAcc ;
_stPathRef.aExecutablePath[0].fDeceleration:=_stSShapedParam.fA_LimDec;

_stPathRef.aExecutablePath[0].fJmax:=_stSShapedParam.fJmax ;
_stPathRef.aExecutablePath[0].fJmin:=_stSShapedParam.fJmin ;

_stPathRef.aExecutablePath[0].fStartPos:=_fStartPos;
_stPathRef.aExecutablePath[0].fEndPos:=_fEndPos;


_stPathRef.bCalculateDone:=TRUE;
stAxis.stAxisStatus.stPathRef:=_stPathRef;
_bCalculateDone:=TRUE;
_fTime:=0;
_nIndex:=0;
stAxis.stAxisStatus.nNcCycleCounter:=0;
END_ACTION

ACTION A_SShapedPosition:
stAxis.stNcTOPLC.nAxisState:=6;
_fTime:=_fTime+fCycleTime;
stAxis.stAxisStatus.nNcCycleCounter:=stAxis.stAxisStatus.nNcCycleCounter+1;


_stAxis_Point:=_fbAxis.M_SShapedPosition(fTime:=_fTime , stS_Parameter:=_stSShapedParam )	;					

//stAxis.stNcTOPLC.fSetPos:=_stAxis_Point.fPosition;
//stAxis.stNcTOPLC.fActPos:=stAxis.stNcTOPLC.fSetPos;
stAxis.stNcTOPLC.fActPos:=_stAxis_Point.fPosition;		
//stAxis.stNcTOPLC.fSetVelo:=_stAxis_Point.fVelocity;  //04.15注释
stAxis.stNcTOPLC.fActVelo:=_stAxis_Point.fVelocity;

IF (_eDirection=E_Direction.DIRECTION_POSITIVE)THEN    //04.15速度方向处理
	 stAxis.stNcTOPLC.fSetVelo:=stAxis.stNcTOPLC.fActVelo;
ELSE
     stAxis.stNcTOPLC.fSetVelo:=-stAxis.stNcTOPLC.fActVelo;
END_IF
	
stAxis.stNcTOPLC.fSetAcc:=_stAxis_Point.fAccleration;  //07.30
stAxis.stNcTOPLC.fSetJerk:=_stAxis_Point.fbJerk;

//stAxis.stNcTOPLC.fModuloSetPos:= ABS(stAxis.stNcTOPLC.fSetPos);
						
// 路径结束条件判断
IF (_fTime>=stAxis.stAxisStatus.stPathRef.aExecutablePath[_nIndex].fTotalTime)THEN
	 _nIndex:=_nIndex+1;
	 _fTime:=0;
	 IF (stAxis.stAxisStatus.stPathRef.aExecutablePath[_nIndex].fTotalTime=0) THEN
	     _fTime:=0;
	     _bCalculateDone:=FALSE;
		 
	     stAxis.stAxisStatus.stPathRef.bCalculateDone:=FALSE;
	     stAxis.stNcTOPLC.nAxisState:=2;
	     stAxis.stAxisStatus.nNcCycleCounter:=0;
		 //stAxis.stNcTOPLC.fSetVelo:=0;
		 stAxis.stNcTOPLC.fActVelo:=0;
	     stAxis.stNcTOPLC.fSetAcc:=0;
		 _fLastPosNC:=0;
		 _nIndex:=0;
		 _bSynMode:=FALSE;
		 //_pPremover^.stAxisStatus.bSynDecActive:=false;
		 stAxis.stAxisStatus.bSynDecActive:=FALSE;
	 END_IF 
END_IF
END_ACTION

ACTION A_StopHandle:

// 增加stop后 后续路径更新功能  根据前动子stop信号停止 01.17
// 不考虑下一段有无动子
IF (stAxis.stAxisStatus.nNcCycleCounter=0)THEN   //03.26
	RETURN;  
END_IF


// 11.04重新梳理逻辑 分为当前动子执行abs指令和fork指令
IF (stAxis.stPLCTONC.nRoadID_1=0) THEN
	IF _pPremover^.stAxisStatus.bSynStopping AND NOT stAxis.stAxisStatus.bSynStopping AND(_pPremover^.stNcTOPLC.nAxisId<>0)THEN //10.28
	   IF (_eDirection=E_Direction.DIRECTION_POSITIVE)THEN
				IF (_pPremover^.stAxisStatus.stPathRef._nPathSegmentNum=1)THEN
					IF (stAxis.stAxisStatus.stPathRef._nPathSegmentNum=1)THEN
						 IF ((_pPremover^.stAxisStatus.stPathRef.aExecutablePath[0].fEndPos-stAxis.stAxisStatus.stPathRef.aExecutablePath[0].fEndPos)<_fGapSet) THEN
							A_UpdateNewTarPos();
							//stAxis.stAxisStatus.bSynStopping:=TRUE;
						 END_IF
					 ELSE
						 IF ((_pPremover^.stAxisStatus.stPathRef.aExecutablePath[0].fEndPos-stAxis.stAxisStatus.stPathRef.aExecutablePath[1].fEndPos)<_fGapSet) THEN
							A_UpdateNewTarPos();
							//stAxis.stAxisStatus.bSynStopping:=TRUE;
						 END_IF
					 END_IF
				ELSE
				    IF (stAxis.stAxisStatus.stPathRef._nPathSegmentNum=1)THEN
					   IF ((_pPremover^.stAxisStatus.stPathRef.aExecutablePath[1].fEndPos-stAxis.stAxisStatus.stPathRef.aExecutablePath[0].fEndPos)<_fGapSet) THEN
					       A_UpdateNewTarPos();
						   //stAxis.stAxisStatus.bSynStopping:=TRUE;
				        END_IF
					ELSE
						IF ((_pPremover^.stAxisStatus.stPathRef.aExecutablePath[1].fEndPos-stAxis.stAxisStatus.stPathRef.aExecutablePath[1].fEndPos)<_fGapSet) THEN
					       A_UpdateNewTarPos();
						  // stAxis.stAxisStatus.bSynStopping:=TRUE;
				        END_IF
					END_IF
				END_IF
	   ELSE
				 IF (_pPremover^.stAxisStatus.stPathRef._nPathSegmentNum=1)THEN
					 IF (stAxis.stAxisStatus.stPathRef._nPathSegmentNum=1)THEN
						   IF ((stAxis.stAxisStatus.stPathRef.aExecutablePath[0].fEndPos-_pPremover^.stAxisStatus.stPathRef.aExecutablePath[0].fEndPos)<_fGapSet)THEN
								
								A_UpdateNewTarPos();
								//stAxis.stAxisStatus.bSynStopping:=TRUE;
						   END_IF
					 ELSE
						 IF ((stAxis.stAxisStatus.stPathRef.aExecutablePath[1].fEndPos-_pPremover^.stAxisStatus.stPathRef.aExecutablePath[0].fEndPos)<_fGapSet)THEN
								
								A_UpdateNewTarPos();
								//stAxis.stAxisStatus.bSynStopping:=TRUE;
						   END_IF
					 END_IF
				 ELSE
					 IF (stAxis.stAxisStatus.stPathRef._nPathSegmentNum=1)THEN
						 IF ((stAxis.stAxisStatus.stPathRef.aExecutablePath[1].fEndPos-_pPremover^.stAxisStatus.stPathRef.aExecutablePath[1].fEndPos)<_fGapSet)
								AND (stAxis.stAxisStatus.stPathRef._nPathSegmentNum=1)  THEN
								A_UpdateNewTarPos();
								//stAxis.stAxisStatus.bSynStopping:=TRUE;
						  END_IF
					 ELSE
						 IF ((stAxis.stAxisStatus.stPathRef.aExecutablePath[1].fEndPos-_pPremover^.stAxisStatus.stPathRef.aExecutablePath[1].fEndPos)<_fGapSet)
								AND (stAxis.stAxisStatus.stPathRef._nPathSegmentNum=1)  THEN
								A_UpdateNewTarPos();
								//stAxis.stAxisStatus.bSynStopping:=TRUE;
						  END_IF
					 END_IF
				 END_IF
	   END_IF 
    END_IF
ELSE  //fork指令 分为当前road和nextroad有无动子 
	IF (_pPremover^.stNcTOPLC.nAxisId<>0) THEN     //前置有动子
		IF (_pPremover^.stPLCTONC.nRoadID_1<>0)AND _pPremover^.stAxisStatus.bSynStopping AND NOT stAxis.stAxisStatus.bSynStopping THEN    //前置动子执行fork指令
			IF (stAxis.stNcTOPLC.nCuRoadID=stAxis.stPLCTONC.nRoadID_1)THEN
				  IF (_eDirection=E_Direction.DIRECTION_POSITIVE)THEN
						IF (_pPremover^.stAxisStatus.stPathRef._nPathSegmentNum=1)THEN
							IF (stAxis.stAxisStatus.stPathRef._nPathSegmentNum=1)THEN
								IF ((_pPremover^.stAxisStatus.stPathRef.aExecutablePath[0].fEndPos-stAxis.stAxisStatus.stPathRef.aExecutablePath[0].fEndPos)<_fGapSet) THEN
									A_UpdateNewTarPos();
									//stAxis.stAxisStatus.bSynStopping:=TRUE;
								END_IF
							ELSE
								IF ((_pPremover^.stAxisStatus.stPathRef.aExecutablePath[0].fEndPos-stAxis.stAxisStatus.stPathRef.aExecutablePath[1].fEndPos)<_fGapSet) THEN
									A_UpdateNewTarPos();
									//stAxis.stAxisStatus.bSynStopping:=TRUE;
								END_IF
							END_IF
						ELSE
							IF (stAxis.stAxisStatus.stPathRef._nPathSegmentNum=1)THEN
								IF ((_pPremover^.stAxisStatus.stPathRef.aExecutablePath[1].fEndPos-stAxis.stAxisStatus.stPathRef.aExecutablePath[0].fEndPos)<_fGapSet) THEN
									A_UpdateNewTarPos();
									//stAxis.stAxisStatus.bSynStopping:=TRUE;
								END_IF	 
                            ELSE
			                    IF ((_pPremover^.stAxisStatus.stPathRef.aExecutablePath[1].fEndPos-stAxis.stAxisStatus.stPathRef.aExecutablePath[1].fEndPos)<_fGapSet) THEN
									A_UpdateNewTarPos();
									//stAxis.stAxisStatus.bSynStopping:=TRUE;
								END_IF
							END_IF 
						END_IF
			      ELSE
						IF (_pPremover^.stAxisStatus.stPathRef._nPathSegmentNum=1)THEN
							IF (stAxis.stAxisStatus.stPathRef._nPathSegmentNum=1)THEN
								IF ((stAxis.stAxisStatus.stPathRef.aExecutablePath[0].fEndPos-_pPremover^.stAxisStatus.stPathRef.aExecutablePath[0].fEndPos)<_fGapSet)THEN
											A_UpdateNewTarPos();
											//stAxis.stAxisStatus.bSynStopping:=TRUE;
								END_IF
							ELSE
								IF ((stAxis.stAxisStatus.stPathRef.aExecutablePath[1].fEndPos-_pPremover^.stAxisStatus.stPathRef.aExecutablePath[0].fEndPos)<_fGapSet)THEN
											A_UpdateNewTarPos();
											//stAxis.stAxisStatus.bSynStopping:=TRUE;
								END_IF
							END_IF
						ELSE
							IF (stAxis.stAxisStatus.stPathRef._nPathSegmentNum=1)THEN
								IF ((stAxis.stAxisStatus.stPathRef.aExecutablePath[0].fEndPos-_pPremover^.stAxisStatus.stPathRef.aExecutablePath[1].fEndPos)<_fGapSet)THEN
										
											A_UpdateNewTarPos();
											//stAxis.stAxisStatus.bSynStopping:=TRUE;
								END_IF
						    ELSE
								IF ((stAxis.stAxisStatus.stPathRef.aExecutablePath[1].fEndPos-_pPremover^.stAxisStatus.stPathRef.aExecutablePath[1].fEndPos)<_fGapSet)THEN
										
											A_UpdateNewTarPos();
											//stAxis.stAxisStatus.bSynStopping:=TRUE;
								END_IF
							END_IF
						END_IF
				  END_IF 
			ELSE
				IF (stAxis.stPLCTONC.stStartPosition.nRoadID=stAxis.stPLCTONC.stEndPosition.nRoadID)THEN 
					IF NOT stAxis.stPLCTONC.bRoadDirection  THEN   //正向 		
								   IF (_pPremover^.stAxisStatus.stPathRef._nPathSegmentNum=1)THEN
									   IF (stAxis.stAxisStatus.stPathRef._nPathSegmentNum=1)THEN
											 IF ((_pPremover^.stAxisStatus.stPathRef.aExecutablePath[0].fEndPos-stAxis.stAxisStatus.stPathRef.aExecutablePath[0].fEndPos)<_fGapSet) THEN
												A_UpdateNewTarPos();
												//stAxis.stAxisStatus.bSynStopping:=TRUE;
											 END_IF
									   ELSE
											 IF ((_pPremover^.stAxisStatus.stPathRef.aExecutablePath[0].fEndPos-stAxis.stAxisStatus.stPathRef.aExecutablePath[1].fEndPos)<_fGapSet) THEN
												A_UpdateNewTarPos();
												//stAxis.stAxisStatus.bSynStopping:=TRUE;
											 END_IF
											
									   END_IF
								   ELSE
									    IF (stAxis.stAxisStatus.stPathRef._nPathSegmentNum=1)THEN
										   IF ((_pPremover^.stAxisStatus.stPathRef.aExecutablePath[1].fEndPos-stAxis.stAxisStatus.stPathRef.aExecutablePath[0].fEndPos)<_fGapSet) THEN
											   A_UpdateNewTarPos();
											   //stAxis.stAxisStatus.bSynStopping:=TRUE;
											END_IF
										ELSE
											IF ((_pPremover^.stAxisStatus.stPathRef.aExecutablePath[1].fEndPos-stAxis.stAxisStatus.stPathRef.aExecutablePath[1].fEndPos)<_fGapSet) THEN
											   A_UpdateNewTarPos();
											   //stAxis.stAxisStatus.bSynStopping:=TRUE;
											END_IF
										END_IF
								   END_IF
				    ELSE
								 IF (_pPremover^.stAxisStatus.stPathRef._nPathSegmentNum=1)THEN
									 IF (stAxis.stAxisStatus.stPathRef._nPathSegmentNum=1)  THEN
										   IF ((stAxis.stAxisStatus.stPathRef.aExecutablePath[0].fEndPos-_pPremover^.stAxisStatus.stPathRef.aExecutablePath[0].fEndPos)<_fGapSet)THEN
												
												A_UpdateNewTarPos();
												//stAxis.stAxisStatus.bSynStopping:=TRUE;  
										   END_IF
									 ELSE
										  IF ((stAxis.stAxisStatus.stPathRef.aExecutablePath[1].fEndPos-_pPremover^.stAxisStatus.stPathRef.aExecutablePath[0].fEndPos)<_fGapSet)THEN
												
												A_UpdateNewTarPos();
												//stAxis.stAxisStatus.bSynStopping:=TRUE;  
										   END_IF
									 END_IF
								 ELSE
									 IF (stAxis.stAxisStatus.stPathRef._nPathSegmentNum=1)  THEN
									     IF ((stAxis.stAxisStatus.stPathRef.aExecutablePath[0].fEndPos-_pPremover^.stAxisStatus.stPathRef.aExecutablePath[1].fEndPos)<_fGapSet)THEN
										
											A_UpdateNewTarPos();
											//stAxis.stAxisStatus.bSynStopping:=TRUE;
									     END_IF 
									 ELSE
										 IF ((stAxis.stAxisStatus.stPathRef.aExecutablePath[1].fEndPos-_pPremover^.stAxisStatus.stPathRef.aExecutablePath[1].fEndPos)<_fGapSet)THEN
										
											A_UpdateNewTarPos();
											//stAxis.stAxisStatus.bSynStopping:=TRUE;
									     END_IF 
									 END_IF
								 END_IF
				    END_IF 
				ELSE
					IF (_eDirection=E_Direction.DIRECTION_POSITIVE)THEN
					      IF NOT stAxis.stPLCTONC.bRoadDirection  THEN   //正向 		
								   IF (_pPremover^.stAxisStatus.stPathRef._nPathSegmentNum=1)THEN
									   IF (stAxis.stAxisStatus.stPathRef._nPathSegmentNum=1)THEN
											 IF ((_pPremover^.stAxisStatus.stPathRef.aExecutablePath[0].fEndPos-stAxis.stAxisStatus.stPathRef.aExecutablePath[0].fEndPos+stAxis.stPLCTONC.fRoad1_Length)<_fGapSet) THEN
												A_UpdateNewTarPos();
												//stAxis.stAxisStatus.bSynStopping:=TRUE;
											 END_IF
									   ELSE
											IF ((_pPremover^.stAxisStatus.stPathRef.aExecutablePath[0].fEndPos-stAxis.stAxisStatus.stPathRef.aExecutablePath[1].fEndPos+stAxis.stPLCTONC.fRoad1_Length)<_fGapSet) THEN
												A_UpdateNewTarPos();
												//stAxis.stAxisStatus.bSynStopping:=TRUE;
											 END_IF
											
									   END_IF
								   ELSE
									    IF (stAxis.stAxisStatus.stPathRef._nPathSegmentNum=1)THEN
										   IF ((_pPremover^.stAxisStatus.stPathRef.aExecutablePath[1].fEndPos-stAxis.stAxisStatus.stPathRef.aExecutablePath[0].fEndPos+stAxis.stPLCTONC.fRoad1_Length)<_fGapSet) THEN
											   A_UpdateNewTarPos();
											  // stAxis.stAxisStatus.bSynStopping:=TRUE;
											END_IF
										ELSE
											IF ((_pPremover^.stAxisStatus.stPathRef.aExecutablePath[1].fEndPos-stAxis.stAxisStatus.stPathRef.aExecutablePath[1].fEndPos+stAxis.stPLCTONC.fRoad1_Length)<_fGapSet) THEN
											   A_UpdateNewTarPos();
											   //stAxis.stAxisStatus.bSynStopping:=TRUE;
											END_IF
										END_IF
								   END_IF
						  ELSE
							   IF (_pPremover^.stAxisStatus.stPathRef._nPathSegmentNum=1)THEN
									   IF (stAxis.stAxisStatus.stPathRef._nPathSegmentNum=1)THEN
											 IF ((stAxis.stPLCTONC.fRoad1_Length+stAxis.stPLCTONC.fRoad2_Length-_pPremover^.stAxisStatus.stPathRef.aExecutablePath[0].fEndPos-stAxis.stAxisStatus.stPathRef.aExecutablePath[0].fEndPos)<_fGapSet) THEN
												A_UpdateNewTarPos();
												//stAxis.stAxisStatus.bSynStopping:=TRUE;
											 END_IF
									   ELSE
											 IF ((stAxis.stPLCTONC.fRoad1_Length+stAxis.stPLCTONC.fRoad2_Length-_pPremover^.stAxisStatus.stPathRef.aExecutablePath[0].fEndPos-stAxis.stAxisStatus.stPathRef.aExecutablePath[1].fEndPos)<_fGapSet) THEN
												A_UpdateNewTarPos();
												//stAxis.stAxisStatus.bSynStopping:=TRUE;
											 END_IF
											
									   END_IF
							   ELSE
									    IF (stAxis.stAxisStatus.stPathRef._nPathSegmentNum=1)THEN
											 IF ((stAxis.stPLCTONC.fRoad1_Length+stAxis.stPLCTONC.fRoad2_Length-_pPremover^.stAxisStatus.stPathRef.aExecutablePath[1].fEndPos-stAxis.stAxisStatus.stPathRef.aExecutablePath[0].fEndPos)<_fGapSet) THEN
												A_UpdateNewTarPos();
												//stAxis.stAxisStatus.bSynStopping:=TRUE;
											 END_IF
									    ELSE
											 IF ((stAxis.stPLCTONC.fRoad1_Length+stAxis.stPLCTONC.fRoad2_Length-_pPremover^.stAxisStatus.stPathRef.aExecutablePath[1].fEndPos-stAxis.stAxisStatus.stPathRef.aExecutablePath[1].fEndPos)<_fGapSet) THEN
												A_UpdateNewTarPos();
												//stAxis.stAxisStatus.bSynStopping:=TRUE;
											 END_IF
											
										END_IF
							   END_IF
						  END_IF
					ELSE
						   IF NOT stAxis.stPLCTONC.bRoadDirection  THEN   //正向 		
								   IF (_pPremover^.stAxisStatus.stPathRef._nPathSegmentNum=1)THEN
									   IF (stAxis.stAxisStatus.stPathRef._nPathSegmentNum=1)THEN
											 IF ((_pPremover^.stAxisStatus.stPathRef.aExecutablePath[0].fEndPos+stAxis.stAxisStatus.stPathRef.aExecutablePath[0].fEndPos)<_fGapSet) THEN
												A_UpdateNewTarPos();
												//stAxis.stAxisStatus.bSynStopping:=TRUE;
											 END_IF
									   ELSE
											IF ((_pPremover^.stAxisStatus.stPathRef.aExecutablePath[0].fEndPos+stAxis.stAxisStatus.stPathRef.aExecutablePath[1].fEndPos)<_fGapSet) THEN
												A_UpdateNewTarPos();
												//stAxis.stAxisStatus.bSynStopping:=TRUE;
											 END_IF
											
									   END_IF
								   ELSE
									    IF (stAxis.stAxisStatus.stPathRef._nPathSegmentNum=1)THEN
										   IF ((_pPremover^.stAxisStatus.stPathRef.aExecutablePath[1].fEndPos+stAxis.stAxisStatus.stPathRef.aExecutablePath[0].fEndPos)<_fGapSet) THEN
											   A_UpdateNewTarPos();
											   //stAxis.stAxisStatus.bSynStopping:=TRUE;
											END_IF
										ELSE
											IF ((_pPremover^.stAxisStatus.stPathRef.aExecutablePath[1].fEndPos+stAxis.stAxisStatus.stPathRef.aExecutablePath[1].fEndPos)<_fGapSet) THEN
											   A_UpdateNewTarPos();
											   //stAxis.stAxisStatus.bSynStopping:=TRUE;
											END_IF
										END_IF
								   END_IF
						   ELSE
							   IF (_pPremover^.stAxisStatus.stPathRef._nPathSegmentNum=1)THEN
									   IF (stAxis.stAxisStatus.stPathRef._nPathSegmentNum=1)THEN
											 IF ((stAxis.stPLCTONC.fRoad2_Length-_pPremover^.stAxisStatus.stPathRef.aExecutablePath[0].fEndPos+stAxis.stAxisStatus.stPathRef.aExecutablePath[0].fEndPos)<_fGapSet) THEN
												A_UpdateNewTarPos();
												//stAxis.stAxisStatus.bSynStopping:=TRUE;
											 END_IF
									   ELSE
											 IF ((stAxis.stPLCTONC.fRoad2_Length-_pPremover^.stAxisStatus.stPathRef.aExecutablePath[0].fEndPos+stAxis.stAxisStatus.stPathRef.aExecutablePath[1].fEndPos)<_fGapSet) THEN
												A_UpdateNewTarPos();
												//stAxis.stAxisStatus.bSynStopping:=TRUE;
											 END_IF
											
									   END_IF
							   ELSE
									    IF (stAxis.stAxisStatus.stPathRef._nPathSegmentNum=1)THEN
											 IF ((stAxis.stPLCTONC.fRoad2_Length-_pPremover^.stAxisStatus.stPathRef.aExecutablePath[1].fEndPos+stAxis.stAxisStatus.stPathRef.aExecutablePath[0].fEndPos)<_fGapSet) THEN
												A_UpdateNewTarPos();
												//stAxis.stAxisStatus.bSynStopping:=TRUE;
											 END_IF
									    ELSE
											 IF ((stAxis.stPLCTONC.fRoad2_Length-_pPremover^.stAxisStatus.stPathRef.aExecutablePath[1].fEndPos+stAxis.stAxisStatus.stPathRef.aExecutablePath[1].fEndPos)<_fGapSet) THEN
												A_UpdateNewTarPos();
												//stAxis.stAxisStatus.bSynStopping:=TRUE;
											 END_IF
										END_IF
							   END_IF
						   END_IF
					END_IF 
				
				END_IF
			END_IF
		ELSE   //前置动子执行abs指令
			IF (_pPremover^.stPLCTONC.nRoadID_1=0)AND _pPremover^.stAxisStatus.bSynStopping AND NOT stAxis.stAxisStatus.bSynStopping THEN
				IF (stAxis.stNcTOPLC.nCuRoadID=stAxis.stPLCTONC.nRoadID_1)THEN   //
						   IF (_eDirection=E_Direction.DIRECTION_POSITIVE)THEN
								IF (_pPremover^.stAxisStatus.stPathRef._nPathSegmentNum=1)THEN
									IF (stAxis.stAxisStatus.stPathRef._nPathSegmentNum=1)THEN
										IF ((_pPremover^.stAxisStatus.stPathRef.aExecutablePath[0].fEndPos-stAxis.stAxisStatus.stPathRef.aExecutablePath[0].fEndPos)<_fGapSet) THEN
											A_UpdateNewTarPos();
											//stAxis.stAxisStatus.bSynStopping:=TRUE;
										END_IF
									ELSE
										IF ((_pPremover^.stAxisStatus.stPathRef.aExecutablePath[0].fEndPos-stAxis.stAxisStatus.stPathRef.aExecutablePath[1].fEndPos)<_fGapSet) THEN
											A_UpdateNewTarPos();
											//stAxis.stAxisStatus.bSynStopping:=TRUE;
										END_IF
									END_IF
								ELSE
									IF (stAxis.stAxisStatus.stPathRef._nPathSegmentNum=1)THEN
										IF ((_pPremover^.stAxisStatus.stPathRef.aExecutablePath[1].fEndPos-stAxis.stAxisStatus.stPathRef.aExecutablePath[0].fEndPos)<_fGapSet) THEN
											A_UpdateNewTarPos();
											//stAxis.stAxisStatus.bSynStopping:=TRUE;
										END_IF	 
									ELSE
										IF ((_pPremover^.stAxisStatus.stPathRef.aExecutablePath[1].fEndPos-stAxis.stAxisStatus.stPathRef.aExecutablePath[1].fEndPos)<_fGapSet) THEN
											A_UpdateNewTarPos();
											//stAxis.stAxisStatus.bSynStopping:=TRUE;
										END_IF
									END_IF 
								END_IF
						   ELSE
								IF (_pPremover^.stAxisStatus.stPathRef._nPathSegmentNum=1)THEN
									IF (stAxis.stAxisStatus.stPathRef._nPathSegmentNum=1)THEN
										IF ((stAxis.stAxisStatus.stPathRef.aExecutablePath[0].fEndPos-_pPremover^.stAxisStatus.stPathRef.aExecutablePath[0].fEndPos)<_fGapSet)THEN
													A_UpdateNewTarPos();
													//stAxis.stAxisStatus.bSynStopping:=TRUE;
										END_IF
									ELSE
										IF ((stAxis.stAxisStatus.stPathRef.aExecutablePath[1].fEndPos-_pPremover^.stAxisStatus.stPathRef.aExecutablePath[0].fEndPos)<_fGapSet)THEN
													A_UpdateNewTarPos();
													//stAxis.stAxisStatus.bSynStopping:=TRUE;
										END_IF
									END_IF
								ELSE
									IF (stAxis.stAxisStatus.stPathRef._nPathSegmentNum=1)THEN
										IF ((stAxis.stAxisStatus.stPathRef.aExecutablePath[0].fEndPos-_pPremover^.stAxisStatus.stPathRef.aExecutablePath[1].fEndPos)<_fGapSet)THEN
												
													A_UpdateNewTarPos();
													//stAxis.stAxisStatus.bSynStopping:=TRUE;
										END_IF
									ELSE
										IF ((stAxis.stAxisStatus.stPathRef.aExecutablePath[1].fEndPos-_pPremover^.stAxisStatus.stPathRef.aExecutablePath[1].fEndPos)<_fGapSet)THEN
												
													A_UpdateNewTarPos();
													//stAxis.stAxisStatus.bSynStopping:=TRUE;
										END_IF
									END_IF
								END_IF
						   END_IF 
				ELSE
						   IF (stAxis.stPLCTONC.stStartPosition.nRoadID=stAxis.stPLCTONC.stEndPosition.nRoadID)THEN 
								IF NOT stAxis.stPLCTONC.bRoadDirection  THEN   //正向 		
											   IF (_pPremover^.stAxisStatus.stPathRef._nPathSegmentNum=1)THEN
												   IF (stAxis.stAxisStatus.stPathRef._nPathSegmentNum=1)THEN
														 IF ((_pPremover^.stAxisStatus.stPathRef.aExecutablePath[0].fEndPos-stAxis.stAxisStatus.stPathRef.aExecutablePath[0].fEndPos)<_fGapSet) THEN
															A_UpdateNewTarPos();
															//stAxis.stAxisStatus.bSynStopping:=TRUE;
														 END_IF
												   ELSE
														IF ((_pPremover^.stAxisStatus.stPathRef.aExecutablePath[0].fEndPos-stAxis.stAxisStatus.stPathRef.aExecutablePath[1].fEndPos)<_fGapSet) THEN
															A_UpdateNewTarPos();
															//stAxis.stAxisStatus.bSynStopping:=TRUE;
														 END_IF
														
													END_IF
											   ELSE
													IF (stAxis.stAxisStatus.stPathRef._nPathSegmentNum=1)THEN
													   IF ((_pPremover^.stAxisStatus.stPathRef.aExecutablePath[1].fEndPos-stAxis.stAxisStatus.stPathRef.aExecutablePath[0].fEndPos)<_fGapSet) THEN
														   A_UpdateNewTarPos();
														   //stAxis.stAxisStatus.bSynStopping:=TRUE;
														END_IF
													ELSE
														IF ((_pPremover^.stAxisStatus.stPathRef.aExecutablePath[1].fEndPos-stAxis.stAxisStatus.stPathRef.aExecutablePath[1].fEndPos)<_fGapSet) THEN
														   A_UpdateNewTarPos();
														   //stAxis.stAxisStatus.bSynStopping:=TRUE;
														END_IF
													END_IF
											   END_IF
								ELSE
											 IF (_pPremover^.stAxisStatus.stPathRef._nPathSegmentNum=1)THEN
												 IF (stAxis.stAxisStatus.stPathRef._nPathSegmentNum=1)  THEN
													   IF ((stAxis.stAxisStatus.stPathRef.aExecutablePath[0].fEndPos-_pPremover^.stAxisStatus.stPathRef.aExecutablePath[0].fEndPos)<_fGapSet)THEN
															
															A_UpdateNewTarPos();
															//stAxis.stAxisStatus.bSynStopping:=TRUE;  
													   END_IF
												  ELSE
													  IF ((stAxis.stAxisStatus.stPathRef.aExecutablePath[1].fEndPos-_pPremover^.stAxisStatus.stPathRef.aExecutablePath[0].fEndPos)<_fGapSet)THEN
															
															A_UpdateNewTarPos();
															//stAxis.stAxisStatus.bSynStopping:=TRUE;  
													   END_IF
												  END_IF
											 ELSE
												 IF (stAxis.stAxisStatus.stPathRef._nPathSegmentNum=1)  THEN
													 IF ((stAxis.stAxisStatus.stPathRef.aExecutablePath[0].fEndPos-_pPremover^.stAxisStatus.stPathRef.aExecutablePath[1].fEndPos)<_fGapSet)THEN
													
														A_UpdateNewTarPos();
														//stAxis.stAxisStatus.bSynStopping:=TRUE;
													 END_IF 
												 ELSE
													 IF ((stAxis.stAxisStatus.stPathRef.aExecutablePath[1].fEndPos-_pPremover^.stAxisStatus.stPathRef.aExecutablePath[1].fEndPos)<_fGapSet)THEN
													
														A_UpdateNewTarPos();
														//stAxis.stAxisStatus.bSynStopping:=TRUE;
													 END_IF 
												 END_IF
											 END_IF
								END_IF 
							ELSE
								IF (_eDirection=E_Direction.DIRECTION_POSITIVE)THEN
									  IF NOT stAxis.stPLCTONC.bRoadDirection  THEN   //正向 		
											   IF (_pPremover^.stAxisStatus.stPathRef._nPathSegmentNum=1)THEN
												   IF (stAxis.stAxisStatus.stPathRef._nPathSegmentNum=1)THEN
														 IF ((_pPremover^.stAxisStatus.stPathRef.aExecutablePath[0].fEndPos-stAxis.stAxisStatus.stPathRef.aExecutablePath[0].fEndPos+stAxis.stPLCTONC.fRoad1_Length)<_fGapSet) THEN
															A_UpdateNewTarPos();
															//stAxis.stAxisStatus.bSynStopping:=TRUE;
														 END_IF
												   ELSE
														IF ((_pPremover^.stAxisStatus.stPathRef.aExecutablePath[0].fEndPos-stAxis.stAxisStatus.stPathRef.aExecutablePath[1].fEndPos+stAxis.stPLCTONC.fRoad1_Length)<_fGapSet) THEN
															A_UpdateNewTarPos();
															//stAxis.stAxisStatus.bSynStopping:=TRUE;
														 END_IF
														
												   END_IF
											   ELSE
													IF (stAxis.stAxisStatus.stPathRef._nPathSegmentNum=1)THEN
													   IF ((_pPremover^.stAxisStatus.stPathRef.aExecutablePath[1].fEndPos-stAxis.stAxisStatus.stPathRef.aExecutablePath[0].fEndPos+stAxis.stPLCTONC.fRoad1_Length)<_fGapSet) THEN
														   A_UpdateNewTarPos();
														  // stAxis.stAxisStatus.bSynStopping:=TRUE;
														END_IF
													ELSE
														IF ((_pPremover^.stAxisStatus.stPathRef.aExecutablePath[1].fEndPos-stAxis.stAxisStatus.stPathRef.aExecutablePath[1].fEndPos+stAxis.stPLCTONC.fRoad1_Length)<_fGapSet) THEN
														   A_UpdateNewTarPos();
														   //stAxis.stAxisStatus.bSynStopping:=TRUE;
														END_IF
													END_IF
											   END_IF
									  ELSE
										   IF (_pPremover^.stAxisStatus.stPathRef._nPathSegmentNum=1)THEN
												    IF (stAxis.stAxisStatus.stPathRef._nPathSegmentNum=1)THEN
														 IF ((stAxis.stPLCTONC.fRoad1_Length+stAxis.stPLCTONC.fRoad2_Length-_pPremover^.stAxisStatus.stPathRef.aExecutablePath[0].fEndPos-stAxis.stAxisStatus.stPathRef.aExecutablePath[0].fEndPos)<_fGapSet) THEN
															A_UpdateNewTarPos();
															//stAxis.stAxisStatus.bSynStopping:=TRUE;
														 END_IF
													ELSE
														 IF ((stAxis.stPLCTONC.fRoad1_Length+stAxis.stPLCTONC.fRoad2_Length-_pPremover^.stAxisStatus.stPathRef.aExecutablePath[0].fEndPos-stAxis.stAxisStatus.stPathRef.aExecutablePath[1].fEndPos)<_fGapSet) THEN
															A_UpdateNewTarPos();
															//stAxis.stAxisStatus.bSynStopping:=TRUE;
														 END_IF
														
													END_IF
										   ELSE
													IF (stAxis.stAxisStatus.stPathRef._nPathSegmentNum=1)THEN
														 IF ((stAxis.stPLCTONC.fRoad1_Length+stAxis.stPLCTONC.fRoad2_Length-_pPremover^.stAxisStatus.stPathRef.aExecutablePath[1].fEndPos-stAxis.stAxisStatus.stPathRef.aExecutablePath[0].fEndPos)<_fGapSet) THEN
															A_UpdateNewTarPos();
															//stAxis.stAxisStatus.bSynStopping:=TRUE;
														 END_IF
													ELSE
														 IF ((stAxis.stPLCTONC.fRoad1_Length+stAxis.stPLCTONC.fRoad2_Length-_pPremover^.stAxisStatus.stPathRef.aExecutablePath[1].fEndPos-stAxis.stAxisStatus.stPathRef.aExecutablePath[1].fEndPos)<_fGapSet) THEN
															A_UpdateNewTarPos();
															//stAxis.stAxisStatus.bSynStopping:=TRUE;
														 END_IF
														
													END_IF
										   END_IF
									  END_IF
								ELSE
									   IF NOT stAxis.stPLCTONC.bRoadDirection  THEN   //正向 		
											   IF (_pPremover^.stAxisStatus.stPathRef._nPathSegmentNum=1)THEN
												   IF (stAxis.stAxisStatus.stPathRef._nPathSegmentNum=1)THEN
														 IF ((_pPremover^.stAxisStatus.stPathRef.aExecutablePath[0].fEndPos+stAxis.stAxisStatus.stPathRef.aExecutablePath[0].fEndPos)<_fGapSet) THEN
															A_UpdateNewTarPos();
													     END_IF
	
												    ELSE
														IF ((_pPremover^.stAxisStatus.stPathRef.aExecutablePath[0].fEndPos+stAxis.stAxisStatus.stPathRef.aExecutablePath[1].fEndPos)<_fGapSet) THEN
															A_UpdateNewTarPos();
															//stAxis.stAxisStatus.bSynStopping:=TRUE;
														END_IF
														
													END_IF
											   ELSE
													IF (stAxis.stAxisStatus.stPathRef._nPathSegmentNum=1)THEN
													   IF ((_pPremover^.stAxisStatus.stPathRef.aExecutablePath[1].fEndPos+stAxis.stAxisStatus.stPathRef.aExecutablePath[0].fEndPos)<_fGapSet) THEN
														   A_UpdateNewTarPos();
														   //stAxis.stAxisStatus.bSynStopping:=TRUE;
														END_IF
													
													ELSE
														IF ((_pPremover^.stAxisStatus.stPathRef.aExecutablePath[1].fEndPos+stAxis.stAxisStatus.stPathRef.aExecutablePath[1].fEndPos)<_fGapSet) THEN
														   A_UpdateNewTarPos();
														   //stAxis.stAxisStatus.bSynStopping:=TRUE;
														END_IF
													END_IF
											   END_IF
									   ELSE
										   IF (_pPremover^.stAxisStatus.stPathRef._nPathSegmentNum=1)THEN
												   IF (stAxis.stAxisStatus.stPathRef._nPathSegmentNum=1)THEN
														 IF ((stAxis.stPLCTONC.fRoad2_Length-_pPremover^.stAxisStatus.stPathRef.aExecutablePath[0].fEndPos+stAxis.stAxisStatus.stPathRef.aExecutablePath[0].fEndPos)<_fGapSet) THEN
															A_UpdateNewTarPos();
															//stAxis.stAxisStatus.bSynStopping:=TRUE;
														 END_IF
												   ELSE
														 IF ((stAxis.stPLCTONC.fRoad2_Length-_pPremover^.stAxisStatus.stPathRef.aExecutablePath[0].fEndPos+stAxis.stAxisStatus.stPathRef.aExecutablePath[1].fEndPos)<_fGapSet) THEN
															A_UpdateNewTarPos();
															//stAxis.stAxisStatus.bSynStopping:=TRUE;
														 END_IF
														
												   END_IF
										   ELSE
													IF (stAxis.stAxisStatus.stPathRef._nPathSegmentNum=1)THEN
														 IF ((stAxis.stPLCTONC.fRoad2_Length-_pPremover^.stAxisStatus.stPathRef.aExecutablePath[1].fEndPos+stAxis.stAxisStatus.stPathRef.aExecutablePath[0].fEndPos)<_fGapSet) THEN
															A_UpdateNewTarPos();
															//stAxis.stAxisStatus.bSynStopping:=TRUE;
														 END_IF
													ELSE
														 IF ((stAxis.stPLCTONC.fRoad2_Length-_pPremover^.stAxisStatus.stPathRef.aExecutablePath[1].fEndPos+stAxis.stAxisStatus.stPathRef.aExecutablePath[1].fEndPos)<_fGapSet) THEN
															A_UpdateNewTarPos();
															//stAxis.stAxisStatus.bSynStopping:=TRUE;
														 END_IF
													END_IF
										   END_IF
									   END_IF
								END_IF 
				            END_IF
				END_IF  
					
				//END_IF
			END_IF
	    END_IF
	ELSE       //nextroad前置有动子 
        //IF (_pNextRoadPremover^.stNcTOPLC.nAxisId<>0)AND (stAxis.stNcTOPLC.nCuRoadID<>_pNextRoadPremover^.stNcTOPLC.nCuRoadID)THEN 
		IF (_pNextRoadPremover^.stNcTOPLC.nAxisId<>0)AND (stAxis.stNcTOPLC.nCuRoadID<>_pNextRoadPremover^.stNcTOPLC.nCuRoadID) 
           AND   _pNextRoadPremover^.stAxisStatus.bSynStopping AND NOT stAxis.stAxisStatus.bSynStopping THEN
             IF (_pNextRoadPremover^.stPLCTONC.stStartPosition.nRoadID<>_pNextRoadPremover^.stPLCTONC.stEndPosition.nRoadID)THEN
				  IF (_pNextRoadPremover^.stPLCTONC.stStartPosition.nRoadID=stAxis.stPLCTONC.stStartPosition.nRoadID)THEN  //起点road相同
					   IF (_eDirection=E_Direction.DIRECTION_POSITIVE)THEN
						   IF ((_pNextRoadPremover^.stAxisStatus.stPathRef.aExecutablePath[0].fEndPos-stAxis.stAxisStatus.stPathRef.aExecutablePath[0].fEndPos)<_fGapSet) THEN
								A_NextPathUpdateNewTarPos();
								//stAxis.stAxisStatus.bSynStopping:=TRUE;
						   END_IF
					   ELSE
						   IF ((stAxis.stAxisStatus.stPathRef.aExecutablePath[0].fEndPos-_pNextRoadPremover^.stAxisStatus.stPathRef.aExecutablePath[0].fEndPos)<_fGapSet)THEN	
								A_NextPathUpdateNewTarPos();
								//stAxis.stAxisStatus.bSynStopping:=TRUE;
						   END_IF
					   END_IF
				  ELSE
					  IF (_eDirection=E_Direction.DIRECTION_POSITIVE)THEN
						   IF NOT stAxis.stPLCTONC.bRoadDirection  THEN
							   IF ((_pNextRoadPremover^.stAxisStatus.stPathRef.aExecutablePath[0].fEndPos+stAxis.stPLCTONC.fRoad1_Length-stAxis.stAxisStatus.stPathRef.aExecutablePath[0].fEndPos)<_fGapSet) THEN
								   A_NextPathUpdateNewTarPos();
								   //stAxis.stAxisStatus.bSynStopping:=TRUE;
						       END_IF
				
						   ELSE
							   IF ((stAxis.stPLCTONC.fRoad2_Length-_pNextRoadPremover^.stAxisStatus.stPathRef.aExecutablePath[0].fEndPos+stAxis.stPLCTONC.fRoad1_Length-stAxis.stAxisStatus.stPathRef.aExecutablePath[0].fEndPos)<_fGapSet) THEN
									A_NextPathUpdateNewTarPos();
									//stAxis.stAxisStatus.bSynStopping:=TRUE;
								END_IF
						   END_IF
					  ELSE
						   IF NOT stAxis.stPLCTONC.bRoadDirection  THEN
								IF ((stAxis.stAxisStatus.stPathRef.aExecutablePath[0].fEndPos+_pNextRoadPremover^.stAxisStatus.stPathRef.aExecutablePath[0].fEndPos)<_fGapSet)THEN		
									A_NextPathUpdateNewTarPos();
									//stAxis.stAxisStatus.bSynStopping:=TRUE;
								END_IF
						   ELSE
								IF ((stAxis.stAxisStatus.stPathRef.aExecutablePath[0].fEndPos+stAxis.stPLCTONC.fRoad2_Length-_pNextRoadPremover^.stAxisStatus.stPathRef.aExecutablePath[0].fEndPos)<_fGapSet)THEN		
									A_NextPathUpdateNewTarPos();
									//stAxis.stAxisStatus.bSynStopping:=TRUE;
								END_IF
							
						   END_IF
					  END_IF
				  END_IF
			 ELSE
					   IF (_eDirection=E_Direction.DIRECTION_POSITIVE)THEN
						   IF NOT stAxis.stPLCTONC.bRoadDirection  THEN
								IF ((_pNextRoadPremover^.stAxisStatus.stPathRef.aExecutablePath[0].fEndPos+stAxis.stPLCTONC.fRoad1_Length-stAxis.stAxisStatus.stPathRef.aExecutablePath[0].fEndPos)<_fGapSet) THEN
									A_NextPathUpdateNewTarPos();
									//stAxis.stAxisStatus.bSynStopping:=TRUE;
								END_IF
						   ELSE
								IF ((stAxis.stPLCTONC.fRoad2_Length-_pNextRoadPremover^.stAxisStatus.stPathRef.aExecutablePath[0].fEndPos+stAxis.stPLCTONC.fRoad1_Length-stAxis.stAxisStatus.stPathRef.aExecutablePath[0].fEndPos)<_fGapSet) THEN
									A_NextPathUpdateNewTarPos();
									//stAxis.stAxisStatus.bSynStopping:=TRUE;
								END_IF
						   END_IF
					   ELSE   //负向
						   IF NOT stAxis.stPLCTONC.bRoadDirection  THEN
								IF ((stAxis.stAxisStatus.stPathRef.aExecutablePath[0].fEndPos+_pNextRoadPremover^.stAxisStatus.stPathRef.aExecutablePath[0].fEndPos)<_fGapSet)THEN		
									A_NextPathUpdateNewTarPos();
									//stAxis.stAxisStatus.bSynStopping:=TRUE;
								END_IF
							ELSE
								IF ((stAxis.stAxisStatus.stPathRef.aExecutablePath[0].fEndPos+stAxis.stPLCTONC.fRoad2_Length-_pNextRoadPremover^.stAxisStatus.stPathRef.aExecutablePath[0].fEndPos)<_fGapSet)THEN		
									A_NextPathUpdateNewTarPos();
									//stAxis.stAxisStatus.bSynStopping:=TRUE;
								END_IF
							
							END_IF
					   END_IF  
			 END_IF
			  
		END_IF
    END_IF   

END_IF


A_EStop();   //04.07注释
END_ACTION

ACTION A_TShaped:
_fStartPos:=stAxis.stNcTOPLC.fActPos;
_stPathRef:=_stNoPathRef;


IF (_fDistance>0)THEN
	_stTimeInfo:=_fbAxis.M_TShaped(
					fVeloStart:=_fVeloStart , 
					fVeloEnd:= _fVeloEnd, 
					fTargetVelo:=_fTargetVelo , 
					fDistance:=_fDistance, 
					fAccleration:=_fAcc , 
					fDeceleration:=_fDec );
ELSE
	RETURN ;
END_IF 

_stPathRef._nPathSegmentNum:=1;
_stPathRef.aExecutablePath[0].fTa:=_stTimeInfo.fTa;
_stPathRef.aExecutablePath[0].fTv:=_stTimeInfo.fTv;
_stPathRef.aExecutablePath[0].fTd:=_stTimeInfo.fTd;
_stPathRef.aExecutablePath[0].fTotalTime:=_stTimeInfo.fT3;
_stPathRef.aExecutablePath[0].fStartVelo:=_fVeloStart;
_stPathRef.aExecutablePath[0].fExpVelo:=_fTargetVelo;
_stPathRef.aExecutablePath[0].fEndVelo:=_fVeloEnd;
_stPathRef.aExecutablePath[0].fAccleration:=_fAcc ;
_stPathRef.aExecutablePath[0].fDeceleration:=_fDec;


_stPathRef.aExecutablePath[0].fStartPos:=_fStartPos;
IF (_eDirection=E_Direction.DIRECTION_POSITIVE)THEN
    _stPathRef.aExecutablePath[0].fEndPos:=_fDistance+_fStartPos;
	_eSetDirection:=E_Direction.DIRECTION_POSITIVE;
	//04.08 终点位置转换
	IF (stAxis.stPLCTONC.nRoadID_1<>0) AND (stAxis.stPLCTONC.nRoadID_2<>0)THEN   
	    IF (stAxis.stPLCTONC.stStartPosition.nRoadID=stAxis.stPLCTONC.nRoadID_2)THEN   
				 IF NOT stAxis.stPLCTONC.bRoadDirection  THEN   //正向 
			         _stPathRef.aExecutablePath[0].fEndPos:=_fDistance+_fStartPos;
					 _eSetDirection:=E_Direction.DIRECTION_POSITIVE;
				 ELSE
					 _stPathRef.aExecutablePath[0].fEndPos:=_fStartPos-_fDistance;
					 _eSetDirection:=E_Direction.DIRECTION_NEGATIVE;
				 END_IF
		 END_IF
	END_IF 
ELSE
	_stPathRef.aExecutablePath[0].fEndPos:=_fStartPos-_fDistance;
	_eSetDirection:=E_Direction.DIRECTION_NEGATIVE;
	//04.28  终点位置转换
	IF (stAxis.stPLCTONC.nRoadID_1<>0) AND (stAxis.stPLCTONC.nRoadID_2<>0)THEN   
	    IF (stAxis.stPLCTONC.stStartPosition.nRoadID=stAxis.stPLCTONC.nRoadID_2)THEN   
				 IF NOT stAxis.stPLCTONC.bRoadDirection  THEN   //正向 
			         _stPathRef.aExecutablePath[0].fEndPos:=_fDistance+_fStartPos;
					 _eSetDirection:=E_Direction.DIRECTION_POSITIVE;
				 ELSE
					 _stPathRef.aExecutablePath[0].fEndPos:=_fStartPos-_fDistance;
					 _eSetDirection:=E_Direction.DIRECTION_NEGATIVE;
				 END_IF
		 END_IF
	END_IF 
END_IF

_stPathRef.aSafePath:=_stPathRef.aExecutablePath;
IF (_eDirection=E_Direction.DIRECTION_POSITIVE)THEN
		
   _stPathRef.aSafePath[0].fStartPos:=_stPathRef.aExecutablePath[0].fStartPos-_fGap;
   _stPathRef.aSafePath[0].fEndPos:=_stPathRef.aExecutablePath[0].fEndPos-_fGap;
   
   //04.08 终点位置转换
	IF (stAxis.stPLCTONC.nRoadID_1<>0) AND (stAxis.stPLCTONC.nRoadID_2<>0)THEN   
	    IF (stAxis.stPLCTONC.stStartPosition.nRoadID=stAxis.stPLCTONC.nRoadID_2)THEN   
				 IF NOT stAxis.stPLCTONC.bRoadDirection  THEN   //正向 
			         _stPathRef.aSafePath[0].fStartPos:=_stPathRef.aExecutablePath[0].fStartPos-_fGap;
                     _stPathRef.aSafePath[0].fEndPos:=_stPathRef.aExecutablePath[0].fEndPos-_fGap;
					 
				 ELSE
					 _stPathRef.aSafePath[0].fStartPos:=_stPathRef.aExecutablePath[0].fStartPos+_fGap;
                      _stPathRef.aSafePath[0].fEndPos:=_stPathRef.aExecutablePath[0].fEndPos+_fGap;
					  
				 END_IF
		 END_IF
	END_IF 
ELSE 
   _stPathRef.aSafePath[0].fStartPos:=_stPathRef.aExecutablePath[0].fStartPos+_fGap;
   _stPathRef.aSafePath[0].fEndPos:=_stPathRef.aExecutablePath[0].fEndPos+_fGap;
   //04.08 终点位置转换
	IF (stAxis.stPLCTONC.nRoadID_1<>0) AND (stAxis.stPLCTONC.nRoadID_2<>0)THEN   
	    IF (stAxis.stPLCTONC.stStartPosition.nRoadID=stAxis.stPLCTONC.nRoadID_2)THEN   
				 IF NOT stAxis.stPLCTONC.bRoadDirection  THEN   //正向 
			         _stPathRef.aSafePath[0].fStartPos:=_stPathRef.aExecutablePath[0].fStartPos-_fGap;
                     _stPathRef.aSafePath[0].fEndPos:=_stPathRef.aExecutablePath[0].fEndPos-_fGap;
					
				 ELSE
					 _stPathRef.aSafePath[0].fStartPos:=_stPathRef.aExecutablePath[0].fStartPos+_fGap;
                      _stPathRef.aSafePath[0].fEndPos:=_stPathRef.aExecutablePath[0].fEndPos+_fGap;
					  
				 END_IF
		 END_IF
	END_IF 
END_IF

_stPathRef.fTargetVelocity:=_fTargetVelo;


IF (_nPathSegment=2)THEN 
	IF (_fDistance_2>0)THEN
		_stTimeInfo_2:=_fbAxis.M_TShaped(
						fVeloStart:=_fVeloStart_2 , 
						fVeloEnd:= _fVeloEnd_2, 
						fTargetVelo:=_fTargetVelo_2 , 
						fDistance:=_fDistance_2, 
						fAccleration:=_fAcc_2 , 
						fDeceleration:=_fDec_2 );
	END_IF 
	
	_stPathRef._nPathSegmentNum:=2;
	_stPathRef.aExecutablePath[1].fTa:=_stTimeInfo_2.fTa;
	_stPathRef.aExecutablePath[1].fTv:=_stTimeInfo_2.fTv;
	_stPathRef.aExecutablePath[1].fTd:=_stTimeInfo_2.fTd;
	_stPathRef.aExecutablePath[1].fTotalTime:=_stTimeInfo_2.fT3;
	_stPathRef.aExecutablePath[1].fStartVelo:=_fVeloStart_2;
	_stPathRef.aExecutablePath[1].fExpVelo:=_fTargetVelo_2;
	_stPathRef.aExecutablePath[1].fEndVelo:= _fVeloEnd_2;
	_stPathRef.aExecutablePath[1].fAccleration:=_fAcc_2 ;
	_stPathRef.aExecutablePath[1].fDeceleration:=_fDec_2;
	_stPathRef.aExecutablePath[1].fStartPos:=_stPathRef.aExecutablePath[0].fEndPos;
	IF (_eDirection=E_Direction.DIRECTION_POSITIVE)THEN
		_stPathRef.aExecutablePath[1].fEndPos:=_fDistance_2+_stPathRef.aExecutablePath[1].fStartPos;
	ELSE
		_stPathRef.aExecutablePath[1].fEndPos:=_stPathRef.aExecutablePath[1].fStartPos-_fDistance_2;
	END_IF
	
	_stPathRef.aSafePath:=_stPathRef.aExecutablePath;
	IF (_eDirection=E_Direction.DIRECTION_POSITIVE)THEN
			
	   _stPathRef.aSafePath[1].fStartPos:=_stPathRef.aExecutablePath[1].fStartPos-_fGap;
	   _stPathRef.aSafePath[1].fEndPos:=_stPathRef.aExecutablePath[1].fEndPos-_fGap;
	ELSE 
	   _stPathRef.aSafePath[1].fStartPos:=_stPathRef.aExecutablePath[1].fStartPos+_fGap;
	   _stPathRef.aSafePath[1].fEndPos:=_stPathRef.aExecutablePath[1].fEndPos+_fGap;
	END_IF
	
	_stPathRef.fTargetVelocity:=_fTargetVelo;
    _stPathRef.fDealtInPos:=  _fPosIn;       //11.29
END_IF
_stPathRef.fGap:=_fGap;
_stPathRef.fSetGap:=stAxis.stAxisStatus.stPathRef.fSetGap;

_stPathRef.bCalculateDone:=TRUE;
stAxis.stAxisStatus.stPathRef:=_stPathRef;

_bCalculateDone:=TRUE;
_fTime:=0;
_nIndex:=0;
stAxis.stAxisStatus.nNcCycleCounter:=0;
IF _bEstopping THEN    //03.03
	stAxis.stAxisStatus.bEmStopping:=TRUE;
END_IF

_stLastAxis_Point.fPosition:=stAxis.stNcTOPLC.fActPos;//03.14

IF GVL_MC.cDebug  THEN
		//_sMessage:=FC_StrContact(stAxis,'NC generate path');
	    // ADSLOGSTR(ADSLOG_MSGTYPE_HINT, _sMessage, '');
	_sMessage2:=FC_StrContactEx(stAxis,'NC cla path');
	 ADSLOGSTR(ADSLOG_MSGTYPE_HINT, _sMessage2, '');
	;	 
END_IF
END_ACTION

ACTION A_TShapedPosition:
 //_nSysType:=stAxis.stPLCTONC.nSysType;   //01.13
 _fRoad1_Lenth:=stAxis.stPLCTONC.fRoad1_Length;
 _fRoad2_Lenth:=stAxis.stPLCTONC.fRoad2_Length;
 
stAxis.stNcTOPLC.nAxisState:=6;
_fTime:=_fTime+fCycleTime;
stAxis.stAxisStatus.nNcCycleCounter:=stAxis.stAxisStatus.nNcCycleCounter+1;

_stAxis_Point:=_fbAxis.M_GetPosition(
						fTime:=_fTime , 
						fTa:=stAxis.stAxisStatus.stPathRef.aExecutablePath[_nIndex].fTa , 
						fTv:=stAxis.stAxisStatus.stPathRef.aExecutablePath[_nIndex].fTv , 
						fTd:=stAxis.stAxisStatus.stPathRef.aExecutablePath[_nIndex].fTd , 
						fVeloStart:=stAxis.stAxisStatus.stPathRef.aExecutablePath[_nIndex].fStartVelo , 
						fVeloEnd:=stAxis.stAxisStatus.stPathRef.aExecutablePath[_nIndex].fEndVelo , 
						fTargetVelo:=stAxis.stAxisStatus.stPathRef.aExecutablePath[_nIndex].fExpVelo , 
						fAccleration:=stAxis.stAxisStatus.stPathRef.aExecutablePath[_nIndex].fAccleration , 
						fDeceleration:=stAxis.stAxisStatus.stPathRef.aExecutablePath[_nIndex].fDeceleration ,   //02.21
						fInitalPos:=stAxis.stAxisStatus.stPathRef.aExecutablePath[_nIndex].fStartPos ,
						eDirection:= _eSetDirection);
						//eDirection:= _eDirection);  //04.08


//  实时位置、速度处理
IF (_nSysType=1)OR(_nSysType=4)	THEN    //接驳线和分叉线
	IF (_eDirection=E_Direction.DIRECTION_POSITIVE)THEN
		IF (stAxis.stPLCTONC.stStartPosition.nRoadID<>stAxis.stPLCTONC.stEndPosition.nRoadID)THEN    //id不相同处理
			IF (_stAxis_Point.fPosition<_fRoad1_Lenth)THEN  //04.16
				//stAxis.stNcTOPLC.fActPos:=floor(_stAxis_Point.fPosition);  //04.19
				stAxis.stNcTOPLC.fActPos:=LTRUNC(_stAxis_Point.fPosition);   //04.19
				stAxis.stNcTOPLC.nCuRoadID:=stAxis.stPLCTONC.nRoadID_1;
			ELSE
				IF NOT stAxis.stPLCTONC.bRoadDirection THEN 
				    stAxis.stNcTOPLC.fActPos:=LTRUNC(FC_TransformPosition(fOffset:=-_fRoad1_Lenth , fPosition:=_stAxis_Point.fPosition ));
				ELSE
					_fPosTemp:=FC_TransformPosition(fOffset:=-_fRoad1_Lenth , fPosition:=_stAxis_Point.fPosition );
					 stAxis.stNcTOPLC.fActPos:= LTRUNC(_fRoad2_Lenth-_fPosTemp);
				END_IF
				
				stAxis.stNcTOPLC.nCuRoadID:=stAxis.stPLCTONC.nRoadID_2;
			END_IF
			stAxis.stNcTOPLC.fSetVelo:=_stAxis_Point.fVelocity;  
			stAxis.stNcTOPLC.fActVelo:=_stAxis_Point.fVelocity;
		ELSE  //ID 相同
			IF (stAxis.stPLCTONC.stEndPosition.nRoadID=stAxis.stPLCTONC.nRoadID_1)THEN   //03.05
			    stAxis.stNcTOPLC.fActPos:=LTRUNC(_stAxis_Point.fPosition);
			    stAxis.stNcTOPLC.nCuRoadID:=stAxis.stPLCTONC.nRoadID_1;
			ELSE 
				
				stAxis.stNcTOPLC.fActPos:=LTRUNC(_stAxis_Point.fPosition);   //04.07
                stAxis.stNcTOPLC.nCuRoadID:=stAxis.stPLCTONC.nRoadID_2;
			END_IF
		    stAxis.stNcTOPLC.fSetVelo:=_stAxis_Point.fVelocity;  
			stAxis.stNcTOPLC.fActVelo:=_stAxis_Point.fVelocity;
		END_IF
	ELSE
		IF (stAxis.stPLCTONC.stStartPosition.nRoadID<>stAxis.stPLCTONC.stEndPosition.nRoadID)THEN    //id不相同处理
			IF (_stAxis_Point.fPosition>0)THEN  //04.16
				stAxis.stNcTOPLC.nCuRoadID:=stAxis.stPLCTONC.nRoadID_1;
				stAxis.stNcTOPLC.fActPos:=LTRUNC(_stAxis_Point.fPosition);
		
			ELSE
				IF NOT stAxis.stPLCTONC.bRoadDirection THEN     //正向
					stAxis.stNcTOPLC.fActPos:=LTRUNC(ABS(_stAxis_Point.fPosition));
				ELSE
					_fPosTemp:=ABS(_stAxis_Point.fPosition);
					stAxis.stNcTOPLC.fActPos:= LTRUNC(_fRoad2_Lenth-_fPosTemp);
				END_IF
				stAxis.stNcTOPLC.nCuRoadID:=stAxis.stPLCTONC.nRoadID_2;
			END_IF
            stAxis.stNcTOPLC.fSetVelo:=_stAxis_Point.fVelocity;  
			stAxis.stNcTOPLC.fActVelo:=_stAxis_Point.fVelocity;
		ELSE
			IF (stAxis.stPLCTONC.stEndPosition.nRoadID=stAxis.stPLCTONC.nRoadID_1)THEN 
				stAxis.stNcTOPLC.fActPos:=LTRUNC(_stAxis_Point.fPosition);
				stAxis.stNcTOPLC.nCuRoadID:=stAxis.stPLCTONC.nRoadID_1;
			ELSE
				stAxis.stNcTOPLC.fActPos:=LTRUNC(_stAxis_Point.fPosition);
                stAxis.stNcTOPLC.nCuRoadID:=stAxis.stPLCTONC.nRoadID_2;
			END_IF
		    stAxis.stNcTOPLC.fSetVelo:=_stAxis_Point.fVelocity;  
			stAxis.stNcTOPLC.fActVelo:=_stAxis_Point.fVelocity;
		END_IF
	
	END_IF
ELSE
    stAxis.stNcTOPLC.fDealtPos:=ABS(LTRUNC(_stAxis_Point.fPosition)-stAxis.stNcTOPLC.fActPos);    //01.13
	stAxis.stNcTOPLC.fActPos:=LTRUNC(_stAxis_Point.fPosition);
	//stAxis.stNcTOPLC.fSetVelo:=floor(_stAxis_Point.fVelocity);  //04.15注释
	stAxis.stNcTOPLC.fActVelo:=LTRUNC(_stAxis_Point.fVelocity);
	IF (_eDirection=E_Direction.DIRECTION_POSITIVE)THEN    //04.15速度方向处理
	    stAxis.stNcTOPLC.fSetVelo:=stAxis.stNcTOPLC.fActVelo;
	ELSE
		stAxis.stNcTOPLC.fSetVelo:=-stAxis.stNcTOPLC.fActVelo;
	END_IF
	
END_IF


// 路径结束条件判断
IF (_fTime>=stAxis.stAxisStatus.stPathRef.aExecutablePath[_nIndex].fTotalTime)THEN
	 _nIndex:=_nIndex+1;
	 _fTime:=0;
	 IF (stAxis.stAxisStatus.stPathRef.aExecutablePath[_nIndex].fTotalTime=0) THEN
	     _fTime:=0;
	     _bCalculateDone:=FALSE;
	     stAxis.stAxisStatus.stPathRef.bCalculateDone:=FALSE;
	     stAxis.stNcTOPLC.nAxisState:=2;
	     stAxis.stAxisStatus.nNcCycleCounter:=0;
		 IF (stAxis.stPLCTONC.stEndPosition.fVelocity=0)THEN   //12.03
		    stAxis.stNcTOPLC.fSetVelo:=0;
		    stAxis.stNcTOPLC.fActVelo:=0;
	         stAxis.stNcTOPLC.fSetAcc:=0;
		 END_IF
		 _fLastPosNC:=0;
		 _nIndex:=0;
		 _bSynMode:=FALSE;
		_bEstopping:=FALSE; //03.19
		 stAxis.stAxisStatus.bSynDecActive:=FALSE;
		 stAxis.stNcTOPLC.fDealtPos:=0;
	 END_IF 
END_IF

 stAxis.stAxisStatus.nSegIndex:=INT_TO_UDINT(_nIndex);
 
 _fLastPtyPos:=stAxis.stCodToNCParam.fActualPos;
END_ACTION

ACTION A_UpdateNewTarPos:
_fAcc:=stAxis.stPLCTONC.stEndPosition.fAccleration;
_fDec:=stAxis.stPLCTONC.stEndPosition.fDeceleration;
//根据指令分类
//IF (stAxis.stPLCTONC.eCommand<>E_Command.COMMAND_ABSOLUTEFORK) THEN	
IF (stAxis.stPLCTONC.nRoadID_1=0)THEN
	IF (_eDirection=E_Direction.DIRECTION_POSITIVE)THEN
		IF (_pPremover^.stAxisStatus.stPathRef._nPathSegmentNum=1)THEN
		    _fUpNewPos:=_pPremover^.stAxisStatus.stPathRef.aExecutablePath[0].fEndPos-_fGapSet-stAxis.stNcTOPLC.fActPos;
		ELSE
			_fUpNewPos:=_pPremover^.stAxisStatus.stPathRef.aExecutablePath[1].fEndPos-_fGapSet-stAxis.stNcTOPLC.fActPos;
		END_IF
	ELSE
		IF (_pPremover^.stAxisStatus.stPathRef._nPathSegmentNum=1)THEN
		    _fUpNewPos:=stAxis.stNcTOPLC.fActPos-_pPremover^.stAxisStatus.stPathRef.aExecutablePath[0].fEndPos-_fGapSet;
		ELSE
			_fUpNewPos:=stAxis.stNcTOPLC.fActPos-_pPremover^.stAxisStatus.stPathRef.aExecutablePath[1].fEndPos-_fGapSet;
		END_IF
	END_IF
ELSE   //fork指令 根据前动子的edpos id 和当前动子roadid分类讨论
	
	IF (_eDirection=E_Direction.DIRECTION_POSITIVE)THEN
		IF (_pPremover^.stAxisStatus.stPathRef._nPathSegmentNum=1)THEN
		    _fUpNewPos:=_pPremover^.stAxisStatus.stPathRef.aExecutablePath[0].fEndPos-_fGapSet-stAxis.stNcTOPLC.fActPos;
		ELSE
			_fUpNewPos:=_pPremover^.stAxisStatus.stPathRef.aExecutablePath[1].fEndPos-_fGapSet-stAxis.stNcTOPLC.fActPos;
		END_IF
	ELSE
		IF (_pPremover^.stAxisStatus.stPathRef._nPathSegmentNum=1)THEN
		    _fUpNewPos:=stAxis.stNcTOPLC.fActPos-_pPremover^.stAxisStatus.stPathRef.aExecutablePath[0].fEndPos-_fGapSet;
		ELSE
			_fUpNewPos:=stAxis.stNcTOPLC.fActPos-_pPremover^.stAxisStatus.stPathRef.aExecutablePath[1].fEndPos-_fGapSet;
		END_IF
	END_IF
     stAxis.stPLCTONC.stStartPosition.nRoadID:=stAxis.stNcTOPLC.nCuRoadID;
	 stAxis.stPLCTONC.stEndPosition.nRoadID:=stAxis.stNcTOPLC.nCuRoadID;
END_IF
	
_fDistance:=_fUpNewPos;
//_fTargetVelo:=stAxis.stNcTOPLC.fActVelo;  //11.1
// 11.01 停止计算距离，根据距离设置目标速度
IF _fDec<>0 THEN  //11.01 
   _fLastPosDeat:=0.5*stAxis.stNcTOPLC.fActVelo*stAxis.stNcTOPLC.fActVelo/_fDec;
END_IF 
IF LTRUNC(_fDistance)<=_fLastPosDeat THEN
	_fTargetVelo:=stAxis.stNcTOPLC.fActVelo;
ELSE
	_fTargetVelo:=stAxis.stPLCTONC.fTargetVelocity;
END_IF

_fVeloStart:=stAxis.stNcTOPLC.fActVelo;
_fVeloEnd:=0;
_bEnable:=TRUE;
_nPathSegment:=1;
stAxis.stAxisStatus.bSynStopping:=TRUE;  //10.28
IF GVL_MC.cDebug  THEN
	_sMessage:=FC_StrContact(stAxis,'SynStoping path');
	 ADSLOGSTR(ADSLOG_MSGTYPE_HINT, _sMessage, '');
END_IF
END_ACTION

END_FUNCTION_BLOCK

(* stored: Version 1.1.0.1, ProductVersion 3.1.4024.12
   POU FTS_NCGenerator: Id {a3e699e1-6dc3-4e5b-87a3-a1da63e6e80a}, SpecialFunc None
   Action A_AccSegmengt: Id {e556f2a2-9616-4837-b2e4-16990e7300f2}
   Action A_CatchUp: Id {25663087-d2e2-40ff-be97-ed1cbef540da}
   Action A_ContantVeloPosition: Id {2a893d99-46b8-4469-b9c6-45731380e179}
   Action A_ConVeloSegment: Id {ce640661-fe09-4246-81be-052f685d7fac}
   Action A_DecSegment: Id {eedab50c-0b0b-432a-8e0d-3f50365d1dd5}
   Action A_DecSegment_2: Id {9171abea-73fd-4d97-9707-eede68f31098}
   Action A_EStop: Id {ca221e54-5765-4fec-ab70-3f1840b84ee4}
   Action A_FollowMasterPlanning: Id {7f355fd4-a936-4c25-8f25-8316de0df815}
   Action A_FollowMaterPosition: Id {9e341724-0b80-4b90-8f95-edc932853870}
   Action A_FollowPlanning: Id {ea6903f6-e733-451c-8ae4-06963fe4de39}
   Action A_FollowPosition: Id {e71e9bd6-7525-4066-98d4-1736a80b95b5}
   Action A_GapControl: Id {9c13e8d5-b985-434e-acac-0d3a380f5b65}
   Action A_GetPosition: Id {d8afa9dd-a313-4b02-a56d-126fac4c918c}
   Action A_LinearPlanning: Id {9739d663-750e-4ea5-815a-5adebacf4a46}
   Action A_LinearPosition: Id {2cb82625-1c0b-4aae-8fd6-db3eed760d9f}
   Action A_NCStartCase: Id {e4c994d2-3844-42d1-be52-39b99b3baa29}
   Action A_NextPathUpdateNewTarPos: Id {3e1f6c41-c875-4756-aa70-7c2dcc0b3de8}
   Action A_NextRoadAccSegmengt: Id {ac652d19-6891-4997-ae37-2b73633fc4a1}
   Action A_NextRoadCatchUp: Id {7c6e550b-30c9-466c-9a74-2323dae631b4}
   Action A_NextRoadConVeloSegment: Id {fa915933-e6c3-4aff-82b0-679c966f5029}
   Action A_NextRoadDecSegment: Id {94fd092d-cd5c-4a9e-8e12-fa6ffeb7db9c}
   Action A_NextRoadDecSegment_2: Id {c482f00a-2b66-4649-9db4-7619faddaaf7}
   Action A_NextRoadGapControl: Id {6650305b-2e4b-4b60-96db-e9bb6a9d8972}
   Action A_NodeConfig: Id {98bb96e2-9143-41c4-870a-0283974cd4c9}
   Action A_NodeUpdate: Id {55b7c2ab-dc1d-49ef-9e01-f8ad29b21658}
   Action A_Planning: Id {54167c9a-5a41-4eb8-bb62-697252ca27a5}
   Action A_Ploynom3Planning: Id {dcfe1d6d-0a14-44aa-8c67-06ee6e411d9f}
   Action A_Ploynom3Position: Id {39384c29-892f-4e67-b4ad-018d035c5fb3}
   Action A_Ploynom5Position: Id {99d591a6-5651-4766-a8d4-7f5693c9e14c}
   Action A_PositionHandle: Id {ed1d1600-9639-4125-9970-1382f471f966}
   Action A_SShapedPlanning: Id {e403a340-83fb-4a79-ab09-98f7d6e97203}
   Action A_SShapedPosition: Id {b6e919a4-ad20-40eb-b16d-787032adac23}
   Action A_StopHandle: Id {57c3d3c2-f95a-421a-8aea-a22c49572d05}
   Action A_TShaped: Id {4139f278-0348-4b3e-b6ec-e75e8e684762}
   Action A_TShapedPosition: Id {45987908-60e2-4541-9d8e-0ee9cc688680}
   Action A_UpdateNewTarPos: Id {224b343e-37bc-49b3-ac49-2b05326ffb6c} *)
